q_stUps.LineInputVoltage_R := i_stState.fInputVoltageRV;
q_stUps.LineInputVoltage_S := i_stState.fInputVoltageSV;
q_stUps.LineInputVoltage_T := i_stState.fInputVoltageTV;
q_stUps.InputFrequency := i_stState.fInputFrequencyHz;
q_stUps.InputCurrent_R := i_stState.fInputCurrentRA;
q_stUps.InputCurrent_S := i_stState.fInputCurrentSA;
q_stUps.InputCurrent_T := i_stState.fInputCurrentTA;
q_stUps.InverterVoltage_R := i_stState.fInverterVoltageRV;
q_stUps.InverterVoltage_S := i_stState.fInverterVoltageSV;
q_stUps.InverterVoltage_T := i_stState.fInverterVoltageTV;
q_stUps.InverterCurrent_R := i_stState.fInverterCurrentRA;
q_stUps.InverterCurrent_S := i_stState.fInverterCurrentSA;
q_stUps.InverterCurrent_T := i_stState.fInverterCurrentTA;
q_stUps.BypassLineVoltage_R := i_stState.fBypassVoltageRV;
q_stUps.BypassLineVoltage_S := i_stState.fBypassVoltageSV;
q_stUps.BypassLineVoltage_T := i_stState.fBypassVoltageTV;
q_stUps.BypassFrequency := i_stState.fBypassFrequencyHz;
q_stUps.LineOutputVoltage_R := i_stState.fOutputVoltageRV;
q_stUps.LineOutputVoltage_S := i_stState.fOutputVoltageSV;
q_stUps.LineOutputVoltage_T := i_stState.fOutputVoltageTV;
q_stUps.FrequencyOutput := i_stState.fOutputFrequencyHz;
q_stUps.OutputCurrent_R := i_stState.fOutputCurrentRA;
q_stUps.OutputCurrent_S := i_stState.fOutputCurrentSA;
q_stUps.OutputCurrent_T := i_stState.fOutputCurrentTA;
q_stUps.DcLinkVoltage := i_stState.fDcLinkVoltageV;
q_stUps.DcLinkVoltage_High := i_stState.fDcLinkHighVoltageV;
q_stUps.DcLinkVoltage_Low := i_stState.fDcLinkLowVoltageV;
q_stUps.BatteryVoltage := i_stState.fBatteryVoltageV;
q_stUps.BatteryCurrent := i_stState.fBatteryCurrentA;
q_stUps.MPI_A_Current := i_stState.fMpiCurrentAA;
q_stUps.MPI_B_Current := i_stState.fMpiCurrentBA;
q_stUps.MPI_C_Current := i_stState.fMpiCurrentCA;
q_stUps.InputApparentPower := i_stState.fInputApparentPowerKva;
q_stUps.OutputApparentPower := i_stState.fOutputApparentPowerKva;
q_stUps.OutputActivePower := i_stState.fOutputActivePowerKw;
q_stUps.Temp1 := i_stState.fTemperature1C;
q_stUps.Temp2 := i_stState.fTemperature2C;
q_stUps.Temp3 := i_stState.fTemperature3C;
q_stUps.Temp4 := i_stState.fTemperature4C;
q_stUps.Temp5 := i_stState.fTemperature5C;
q_stUps.Temp6 := i_stState.fBatteryRoomTemperatureC;

END_FUNCTION_BLOCK

// ---- 20_Module/Report/FB_RptLsImd1000.TcPOU
FUNCTION_BLOCK FB_RptLsImd1000		// LS IMD1000 읽은 값 → IMD 보고값 (인터페이스\22. IMD.xlsx)
(* 2026-11-09. 명세 DV-11·RD-IMD-01 (v1.8)
   Status (사용자 결정 2026-11-09, 저항이 높은 경보부터)
     b0 통신에러 = 통신 이상 또는 아직 못 읽음 (나머지 칸 0)
     b1 Pre-Warning = Pre Alarm#3 동작 (IR 210 b3, 초기값 100 kΩ)
     b2 Warning = Pre Alarm#1 OR #2 동작 (IR 210 b1·b2, 초기값 40·70 kΩ)
     b3 Fault = 자가진단 오류 (IR 209 b0~2 메모리·RTC·교정) OR Device 이상 (IR 211 b1)
     b4 Alarm = Ins. Alarm 동작 (IR 210 b0, 초기값 10 kΩ)
     b5 Internal test = Self Test 진행 중 (IR 215 = 1)
     b6 External test = 버튼·DI Self Test 입력 (IR 206 b0·b1)
   Fault1 b0 = System 연결 이상 (IR 211 b2), b1 = PE 연결 이상 (IR 211 b0)
   PreAlarmSettingValue = Pre Alarm#1 Pick-up, MainAlarmSettingValue = Ins. Alarm Pick-up (설정 영역을 못 읽었으면 0)
   DeviceErrorLocation·InsulationResistanceFaultLocation은 Bender 항목이라 0 *)
VAR_INPUT
	i_stState		: ST_LsImd1000State;	// 장비 상태 (FB_LsImd1000.q_stState)
	i_nDeviceIndex	: UDINT;				// IMD 번호 (1부터)
END_VAR
VAR_OUTPUT
	q_stImd			: ST_ImdPublish_V1;		// IMD 보고값
	q_bValid		: BOOL;					// 유효한 장비 데이터
END_VAR
VAR
	_stEmpty		: ST_ImdPublish_V1;
END_VAR

q_stImd := _stEmpty;
q_stImd.DeviceIndex := i_nDeviceIndex;
q_stImd.Status := 1;	// b0 통신에러
q_bValid := i_stState.bValid;
IF NOT q_bValid THEN
	RETURN;
END_IF

q_stImd.Status := 0;
q_stImd.Status.1 := i_stState.wAlarm.3;
q_stImd.Status.2 := i_stState.wAlarm.1 OR i_stState.wAlarm.2;
q_stImd.Status.3 := (i_stState.wSelfDiag AND 16#0007) <> 0 OR i_stState.wConnect.1;
q_stImd.Status.4 := i_stState.wAlarm.0;
q_stImd.Status.5 := i_stState.wSelfTest = 1;
q_stImd.Status.6 := i_stState.wDiState.0 OR i_stState.wDiState.1;

q_stImd.InsulationResistance := i_stState.fInsulation;
IF i_stState.bSetValid THEN
	q_stImd.PreAlarmSettingValue := i_stState.nPre1Pickup;
	q_stImd.MainAlarmSettingValue := i_stState.nInsPickup;
END_IF
q_stImd.Fault1.0 := i_stState.wConnect.2;
q_stImd.Fault1.1 := i_stState.wConnect.0;

END_FUNCTION_BLOCK

// ---- 20_Module/Report/FB_RptTempHum.TcPOU
FUNCTION_BLOCK FB_RptTempHum		// 온습도계 읽은 값 → 온도 보고값 (인터페이스\07.Temperature Sensor.xlsx, 토픽 temperature_sensor)
(* 2026-11-09. status b0 통신에러(통신 이상·값 무효면 1, 온도·습도 0). location은 설치 위치 번호
   (1 PCS실, 2 BAT실, 3 UPS실, 4 FC 컨테이너실, 5 외부) *)
VAR_INPUT
	i_stState		: ST_TempHumState;		// 장비 상태 (드라이버 q_stState)
	i_nDeviceIndex	: UDINT;				// 장치 번호 (0부터, 기존 temperature_sensor 시험 데이터와 같음)
	i_nLocation		: UDINT;				// 설치 위치
END_VAR
VAR_OUTPUT
	q_stTemp		: ST_TempPublish_V1;	// 보고값
	q_bValid		: BOOL;					// 유효한 장비 데이터
END_VAR
VAR
	_stEmpty		: ST_TempPublish_V1;
END_VAR

q_stTemp := _stEmpty;
q_stTemp.DeviceIndex := i_nDeviceIndex;
q_stTemp.location := i_nLocation;
q_stTemp.status := 1;	// b0 통신에러
q_bValid := i_stState.bValid;
IF NOT q_bValid THEN
	RETURN;
END_IF
q_stTemp.status := 0;
q_stTemp.temperature := i_stState.fTemp;
q_stTemp.humidity := i_stState.fHum;

END_FUNCTION_BLOCK

// ---- 20_Module/Driver/Esolution/FB_BmsRackCommand.TcPOU
FUNCTION_BLOCK FB_BmsRackCommand		// BMS 랙 컨택터 개별 제어: EMS 랙 명령 → 랙 선택표(BMS 40001 랙 비트) 갱신 요청
(* 2026-11-10. 명세 WR-BAT-01 (v2.5). 인터페이스 100.Command BAT CommandType 11 랙 닫기 / 12 랙 열기 (Value = 랙 번호)
   BAT 질의 Q4 답변: 랙 개별·일괄 제어 모두 지원. 일괄은 CommandType 1·2 (시스템 컨택터 40013, 기존 코어 경로)
   - 랙 선택표(비트 n-1 = 랙 n, 1 = 사용)를 기억하고, 명령마다 그 랙 비트만 바꾼 표 전체를 BMS에 쓰게 한다
   - 장비 쓰기는 하지 않는다. q_bWriteReq·q_wWriteMask를 MAIN이 보고 드라이버 M_SetRackMask를 부르고 결과를 돌려준다
   - 선택표는 PERSISTENT (i_wRestore로 시작 때 한 번 읽고, q_wMask를 MAIN이 저장). 저장값이 없으면(0) 설치된 랙 전부
   - 거절: 랙 번호 범위 밖(BadRequest), 마지막 남은 랙 열기(BadRequest: 0이면 BMS가 전 랙 사용 안 함 → 전체는 일괄 2 열기로)
   - 드라이버가 바쁘면(Busy) WRITE_TIMEOUT 동안 다시 시도. 그 밖의 거절(쓰기 막힘, 통신 불가 등)은 바로 그 결과로 끝
   - 같은 상태로 바꾸는 명령도 표 전체를 다시 씀 (BMS가 다시 켜져 표가 달라졌을 때 맞춤)
   - [2026-11-13] BMS 맵 v1.4 랙 컨택터 상태(Input 30027)를 받으면 그 실제 상태를 바탕으로 비트를 바꿈.
     40013(랙 전체 연결)으로 다 붙은 뒤 옛 선택표로 써서 다른 랙을 떼는 일을 막음. 상태가 없으면 기억한 선택표 *)
VAR_INPUT
	i_stCmd			: ST_BatRackCmd;	// EMS 랙 명령 (번호가 바뀌면 새 명령)
	i_nRackCount	: UINT;				// 설치된 랙 수 (GVL_PARAM.RACKS_PER_BMS)
	i_wRestore		: WORD;				// 처음 호출 때 한 번 읽는 저장된 선택표 (GVL_PERSIST.g_awBmsRackMask[n])
	i_bAccepted		: BOOL;				// 지난 스캔의 쓰기 요청을 드라이버가 받음 (M_SetRackMask 반환값)
	i_eDriverResult	: E_UpsResult;		// 지난 스캔 드라이버 결과 (q_eRequestResult). 요청하지 않은 스캔은 None
	i_wActual		: WORD;				// BMS 랙 컨택터 실제 상태 (q_stState.wRackContactor, 30027) [2026-11-13]
	i_bActualValid	: BOOL;				// i_wActual을 믿을 수 있음 (q_stState.bContactorFeedbackKnown)
END_VAR
VAR_OUTPUT
	q_wMask			: WORD;				// 지금 선택표 (드라이버가 받은 값). MAIN이 GVL_PERSIST에 씀
	q_bMaskChanged	: BOOL;				// 이 스캔에 q_wMask가 바뀜 (PERSISTENT 바로 저장 요청)
	q_bWriteReq		: BOOL;				// 드라이버에 쓰기 요청 중
	q_wWriteMask	: WORD;				// 쓸 선택표
	q_eResult		: E_UpsResult;		// 마지막 명령 결과
	q_nLastSeq		: UDINT;			// 마지막으로 처리한 명령 번호
END_VAR
VAR
	_bInit			: BOOL;
	_wInstalled		: WORD;
	_wNew			: WORD;
	_wOld			: WORD;
	_wBase			: WORD;				// 바꿀 바탕 (실제 상태 또는 기억한 선택표)
	_tonWait		: TON;
END_VAR
VAR CONSTANT
	WRITE_TIMEOUT	: TIME := T#5S;		// 드라이버가 바쁠 때 다시 시도하는 시간
END_VAR

q_bMaskChanged := FALSE;
_wInstalled := SHL(WORD#1, MIN(i_nRackCount, 16)) - 1;
IF NOT _bInit THEN
	q_wMask := i_wRestore AND _wInstalled;
	IF q_wMask = 0 THEN
		q_wMask := _wInstalled;	// 저장값 없음 → 설치된 랙 전부
	END_IF
	_bInit := TRUE;
END_IF
_wOld := q_wMask;

// 1) 지난 스캔 쓰기 요청의 결과
IF q_bWriteReq THEN
	_tonWait(IN := TRUE, PT := WRITE_TIMEOUT);
	IF i_bAccepted THEN
		q_wMask := q_wWriteMask;
		q_eResult := E_UpsResult.Accepted;
		q_bWriteReq := FALSE;
	ELSIF i_eDriverResult <> E_UpsResult.None AND i_eDriverResult <> E_UpsResult.Busy THEN
		q_eResult := i_eDriverResult;	// 쓰기 막힘, 통신 불가, 설정 오류 등
		q_bWriteReq := FALSE;
	ELSIF _tonWait.Q THEN
		q_eResult := E_UpsResult.Busy;	// 계속 바빠서 포기
		q_bWriteReq := FALSE;
	END_IF
	IF NOT q_bWriteReq THEN
		_tonWait(IN := FALSE);
	END_IF
END_IF

// 2) 새 명령 (처리 중인 요청이 있으면 그것을 버리고 새 명령으로)
IF i_stCmd.nSeq <> q_nLastSeq AND i_stCmd.nSeq <> 0 THEN
	q_nLastSeq := i_stCmd.nSeq;
	q_bWriteReq := FALSE;
	_tonWait(IN := FALSE);
	IF i_stCmd.nRack < 1 OR i_stCmd.nRack > i_nRackCount OR i_stCmd.nRack > 16 THEN
		q_eResult := E_UpsResult.BadRequest;
	ELSE
		IF i_bActualValid THEN
			_wBase := i_wActual AND _wInstalled;	// 실제 상태 바탕
		ELSE
			_wBase := q_wMask;
		END_IF
		IF i_stCmd.bClose THEN
			_wNew := _wBase OR SHL(WORD#1, i_stCmd.nRack - 1);
		ELSE
			_wNew := _wBase AND NOT SHL(WORD#1, i_stCmd.nRack - 1);
		END_IF
		IF _wNew = 0 THEN
			q_eResult := E_UpsResult.BadRequest;	// 마지막 랙: 전체 열기는 일괄 명령(2)으로
		ELSE
			q_wWriteMask := _wNew;
			q_bWriteReq := TRUE;
			q_eResult := E_UpsResult.None;	// 처리 중
		END_IF
	END_IF
END_IF

q_bMaskChanged := q_wMask <> _wOld;

END_FUNCTION_BLOCK

// ---- 20_Module/Driver/Esolution/FB_BmsContactorCommand.TcPOU
FUNCTION_BLOCK FB_BmsContactorCommand		// BMS 컨택터 하나씩 제어: EMS 명령 번호 5~10 → 드라이버 M_SetControl 요청
(* 2026-11-13. 인터페이스 100.Command BAT CommandType 5~10, BMS 맵 v1.4 Holding 40013~40015
   5 시스템(랙 전체 40013) 연결   6 시스템 차단
   7 충전 컨택터(40014) 닫기      8 충전 컨택터 열기
   9 방전 컨택터(40015) 닫기      10 방전 컨택터 열기
   - 장비 쓰기는 하지 않는다. q_bWriteReq·q_eControl·q_bOn을 MAIN이 보고 드라이버 M_SetControl을 부르고 결과를 돌려준다
   - 5~10 밖이면 BadRequest. 드라이버가 바쁘면(Busy) WRITE_TIMEOUT 동안 다시 시도. 그 밖의 거절(쓰기 막힘, 통신 불가 등)은 바로 그 결과로 끝
   - 코어 순서(유닛 정지 확인)는 거치지 않는다 (랙 개별 11·12와 같음). 일괄 투입·개방은 1·2 (코어 경로) *)
VAR_INPUT
	i_stCmd			: ST_BatCtlCmd;		// EMS 명령 (번호가 바뀌면 새 명령)
	i_bAccepted		: BOOL;				// 지난 스캔의 쓰기 요청을 드라이버가 받음 (M_SetControl 반환값)
	i_eDriverResult	: E_UpsResult;		// 지난 스캔 드라이버 결과 (q_eRequestResult). 요청하지 않은 스캔은 None
END_VAR
VAR_OUTPUT
	q_bWriteReq		: BOOL;				// 드라이버에 쓰기 요청 중
	q_eControl		: E_EsolutionControl;	// 쓸 컨택터
	q_bOn			: BOOL;				// TRUE = 닫기(붙이기), FALSE = 열기(떼기)
	q_eResult		: E_UpsResult;		// 마지막 명령 결과
	q_nLastSeq		: UDINT;			// 마지막으로 처리한 명령 번호
END_VAR
VAR
	_tonWait		: TON;
END_VAR
VAR CONSTANT
	WRITE_TIMEOUT	: TIME := T#5S;		// 드라이버가 바쁠 때 다시 시도하는 시간
END_VAR

// 1) 지난 스캔 쓰기 요청의 결과
IF q_bWriteReq THEN
	_tonWait(IN := TRUE, PT := WRITE_TIMEOUT);
	IF i_bAccepted THEN
		q_eResult := E_UpsResult.Accepted;
		q_bWriteReq := FALSE;
	ELSIF i_eDriverResult <> E_UpsResult.None AND i_eDriverResult <> E_UpsResult.Busy THEN
		q_eResult := i_eDriverResult;	// 쓰기 막힘, 통신 불가 등
		q_bWriteReq := FALSE;
	ELSIF _tonWait.Q THEN
		q_eResult := E_UpsResult.Busy;	// 계속 바빠서 포기
		q_bWriteReq := FALSE;
	END_IF
	IF NOT q_bWriteReq THEN
		_tonWait(IN := FALSE);
	END_IF
END_IF

// 2) 새 명령 (처리 중인 요청이 있으면 그것을 버리고 새 명령으로)
IF i_stCmd.nSeq <> q_nLastSeq AND i_stCmd.nSeq <> 0 THEN
	q_nLastSeq := i_stCmd.nSeq;
	q_bWriteReq := FALSE;
	_tonWait(IN := FALSE);
	q_eResult := E_UpsResult.None;	// 처리 중
	CASE i_stCmd.nType OF
		5, 6:	q_eControl := E_EsolutionControl.SystemContactor;
		7, 8:	q_eControl := E_EsolutionControl.ChargeContactor;
		9, 10:	q_eControl := E_EsolutionControl.DischargeContactor;
	ELSE
		q_eResult := E_UpsResult.BadRequest;
	END_CASE
	IF q_eResult = E_UpsResult.None THEN
		q_bOn := (i_stCmd.nType MOD 2) = 1;	// 5·7·9 = 닫기
		q_bWriteReq := TRUE;
	END_IF
END_IF

END_FUNCTION_BLOCK

// ---- 20_Module/Ups/FB_UpsSafetyStage.TcPOU
(* LiB-UPS 사고·고장 단계 판정 (④보호 표시 / 장치: UPS·BAT). 2026-11-05.
   기반 없음(신규). 동작시퀀스 7쪽(이솔루션 2026-10-23) 단계표를 따른다.
   변경: 2026-11-09 UPS 경고·고장 4번 칸을 없앰. STATUS 비트를 Warning3 하위·Fault3 상위에서 읽음 (명세 RD-UPS-02 v1.6)
   부호·단위: 해당 없음. 명세: C:\gil\UPS\명세서\UPS_명세서.md SQ-01, WR-SQ-01
   차단·정지는 UPS(UMS)와 BMS가 스스로 한다. 이 FB는 판정과 표시만 하고 장비에 아무것도 쓰지 않는다. *)
FUNCTION_BLOCK FB_UpsSafetyStage
VAR_INPUT
	i_stUps			: ST_UpsPublish_V1;	// UPS 보고값 (FB_RptSebangUps.q_stUps)
	i_bUpsValid		: BOOL;				// UPS 데이터 유효 (통신 정상)
	i_stBat			: ST_BatPublish_V1;	// 짝 BAT 보고값 (FB_RptEsolutionBat.q_stBat)
	i_bBatValid		: BOOL;				// BAT 데이터 유효 (통신 정상)
	i_bAck			: BOOL;				// Fault 단계 확인 (상승 에지). 원인이 해소된 Fault 표시만 내린다 (WR-SQ-01)
END_VAR
VAR_OUTPUT
	q_nStage		: UINT;				// 대표 단계 0~6 (걸린 단계 중 가장 높은 것)
	q_wStageMask	: WORD;				// 걸린 단계 목록. bit n = n단계 (n = 1~6). 높은 순서로 모두 표시할 때 사용
	q_nCause		: UDINT;			// 원인 비트 (아래 CAUSE_* 표). 지금 걸린 원인 + 확인 전인 Fault 원인
	q_nActiveCause	: UDINT;			// 지금 실제로 걸린 원인만
	q_bAckPending	: BOOL;				// 원인은 해소됐지만 운영자 확인 전인 Fault 원인이 있음
	q_bUpsCommFault	: BOOL;				// UPS 통신장애 (단계와 별도 상태). 끊긴 동안 UPS 원인은 마지막 값을 유지
	q_bBatCommFault	: BOOL;				// BAT 통신장애 (단계와 별도 상태). 끊긴 동안 BAT 원인은 마지막 값을 유지
END_VAR
VAR
	_rtAck			: R_TRIG;
	_nUpsCause		: UDINT;			// UPS에서 나온 원인 (통신이 끊기면 마지막 값 유지)
	_nBatCause		: UDINT;			// BAT에서 나온 원인 (통신이 끊기면 마지막 값 유지)
	_nLatched		: UDINT;			// 확인 전까지 유지하는 Fault 원인
	_i				: INT;
END_VAR
VAR CONSTANT
	(* 원인 비트 → 단계. 순서 = 비트 번호 *)
	CAUSE_STAGE		: ARRAY[0..12] OF UINT := [
		1,	// b0  AC·DC SPD (I51 b8·b9)
		1,	// b1  UPS 경고장 (SPD·BMS Minor 제외)
		2,	// b2  BMS Minor (I51 b10)
		3,	// b3  BMS Major (I51 b11)
		3,	// b4  UPS 입력·정류부 중고장 (Fault1)
		3,	// b5  UPS 출력 중고장 (Fault2 상위)
		3,	// b6  UPS 인버터 중고장 (Fault3 하위)
		3,	// b7  배터리 DC 전로 지락 1단계 = RCD 1단계 (I51 b12, 추정)
		4,	// b8  배터리 컨버터(BBC) 중고장 (Fault2 하위)
		4,	// b9  지락 2단계 = RCD 2단계 (I51 b13, 추정)
		5,	// b10 BMS Level 3 (BAT Status b9 System Lock)
		5,	// b11 화재 (I51 b14)
		6];	// b12 ESD (I50 b0)
	FAULT_CAUSE_MASK : UDINT := 16#00001F00;	// 4~6단계 원인 (b8~b12): 확인 전까지 유지
	(* UPS 보고 칸 안의 비트 (명세 RD-UPS-02 v1.6). Warning3 하위 16비트 = I51 경고, Fault3 상위 16비트 = I50 고장 OR I51 고장 *)
	W3_SPD			: UDINT := 16#00000300;	// Warning3: I51 b8 AC SPD, b9 DC SPD
	W3_BMS_MINOR	: UDINT := 16#00000400;	// Warning3: I51 b10
	F3_BMS_MAJOR	: UDINT := 16#08000000;	// Fault3: I51 b11
	F3_RCD1			: UDINT := 16#10000000;	// Fault3: I51 b12
	F3_RCD2			: UDINT := 16#20000000;	// Fault3: I51 b13
	F3_FIRE			: UDINT := 16#40000000;	// Fault3: I51 b14
	F3_ESD			: UDINT := 16#00010000;	// Fault3: I50 b0
	LOWER_WORD		: UDINT := 16#0000FFFF;
	UPPER_WORD		: UDINT := 16#FFFF0000;
END_VAR

// 1) UPS 원인. 통신이 끊기면 마지막 값을 그대로 둔다 (단계를 내리지 않음)
q_bUpsCommFault := NOT i_bUpsValid;
IF i_bUpsValid THEN
	_nUpsCause := 0;
	IF (i_stUps.Warning3 AND W3_SPD) <> 0 THEN _nUpsCause := _nUpsCause OR 16#0001; END_IF
	IF (i_stUps.Warning1 OR i_stUps.Warning2 OR (i_stUps.Warning3 AND NOT (W3_SPD OR W3_BMS_MINOR))) <> 0 THEN _nUpsCause := _nUpsCause OR 16#0002; END_IF
	IF (i_stUps.Warning3 AND W3_BMS_MINOR) <> 0 THEN _nUpsCause := _nUpsCause OR 16#0004; END_IF
	IF (i_stUps.Fault3 AND F3_BMS_MAJOR) <> 0 THEN _nUpsCause := _nUpsCause OR 16#0008; END_IF
	IF i_stUps.Fault1 <> 0 THEN _nUpsCause := _nUpsCause OR 16#0010; END_IF
	IF (i_stUps.Fault2 AND UPPER_WORD) <> 0 THEN _nUpsCause := _nUpsCause OR 16#0020; END_IF
	IF (i_stUps.Fault3 AND LOWER_WORD) <> 0 THEN _nUpsCause := _nUpsCause OR 16#0040; END_IF
	IF (i_stUps.Fault3 AND F3_RCD1) <> 0 THEN _nUpsCause := _nUpsCause OR 16#0080; END_IF
	IF (i_stUps.Fault2 AND LOWER_WORD) <> 0 THEN _nUpsCause := _nUpsCause OR 16#0100; END_IF
	IF (i_stUps.Fault3 AND F3_RCD2) <> 0 THEN _nUpsCause := _nUpsCause OR 16#0200; END_IF
	IF (i_stUps.Fault3 AND F3_FIRE) <> 0 THEN _nUpsCause := _nUpsCause OR 16#0800; END_IF
	IF (i_stUps.Fault3 AND F3_ESD) <> 0 THEN _nUpsCause := _nUpsCause OR 16#1000; END_IF
END_IF

// 2) BAT 원인
q_bBatCommFault := NOT i_bBatValid;
IF i_bBatValid THEN
	_nBatCause := 0;
	IF i_stBat.Status.9 THEN _nBatCause := _nBatCause OR 16#0400; END_IF	// BMS Level 3 (System Lock)
END_IF

q_nActiveCause := _nUpsCause OR _nBatCause;

// 3) Fault(4~6단계)는 원인이 사라져도 확인 전까지 유지. 확인하면 해소된 것만 내림
_nLatched := _nLatched OR (q_nActiveCause AND FAULT_CAUSE_MASK);
_rtAck(CLK := i_bAck);
IF _rtAck.Q THEN
	_nLatched := _nLatched AND q_nActiveCause;
END_IF
q_nCause := q_nActiveCause OR _nLatched;
q_bAckPending := (_nLatched AND NOT q_nActiveCause) <> 0;

// 4) 단계 목록과 대표 단계
q_wStageMask := 0;
q_nStage := 0;
FOR _i := 0 TO 12 DO
	IF (q_nCause AND SHL(UDINT#1, _i)) <> 0 THEN
		q_wStageMask := q_wStageMask OR SHL(WORD#1, CAUSE_STAGE[_i]);
		q_nStage := MAX(q_nStage, CAUSE_STAGE[_i]);
	END_IF
END_FOR

END_FUNCTION_BLOCK

// ---- 20_Module/Mqtt/FB_EmsConfigApply.TcPOU
FUNCTION_BLOCK FB_EmsConfigApply		// EMS config(pcs·bat) → 운영 설정 (PlcTask. MAIN 액션 A_PassEmsCfg가 부름) [9-21 수정 2026-11-04: 추가]
(* - 입력 i_stCfg는 MAIN이 GVL_IF.g_stEmsCfg에서 일관되게 복사해 넘김. PCS·BMS 칸마다 번호(anPcsSeq·anBatSeq)가 바뀌면 새 레코드
   - [21번 수정 2026-11-09] is_available = 0인 값은 기본값으로 반영 (원래: 바꾸지 않고 기존 값 유지 → EMS가 한도를 풀 수 없었음)
       pcs 충전·방전 한도 0 → 그 방향 정격 (= 제한 없음). 두 방향 모두 0 → 그 PCS 유닛의 사용자 P 한도 끔 (bPEnable FALSE, 값은 ±정격)
       bat SOC 하한 0 → 0 %, 상한 0 → 100 % (감발 폭 fBand·재개 마진은 HMI 설정 그대로)
   - [UPS 2026-11-10] UPS 현장의 config/bat 레코드는 103.Config BAT UPS_V1 형식 (SocMin·SocMax = REAL, is_available 없음. UPS_MQTT_INTERFACE.md).
       그래서 bat 값은 받은 BMS(_abBatRx)만 계산에 넣고 항상 '있음'으로 봄. 아직 못 받은 BMS는 기본값(0 %·100 %)과 같아 결과에 영향 없음. pcs 쪽은 STD 그대로
   - pcs: 충전·방전 전력 한도 (kW) → 사용자 한도 stUnitLimit. 그 PCS의 유닛들에 정격 비율로 나눔, 충전은 fPMin (−). PvMarginRate는 쓰지 않음 (사양 대기)
   - bat: SOC 최소·최대 (%) → SOC 정책 stSocLimit. 배터리 그룹 전체 한 세트라 받은 BMS 값(기본값 포함) 중 가장 엄격한 값 (하한 = 가장 큰 값, 상한 = 가장 작은 값)
   - 범위 검사를 먼저 하고 통과한 값만 씀 (SOC는 FB_SocLimit.M_CheckSet과 같은 F_SocLimitSetErr). 버리면 q_bRejected (이벤트 로그 '잘못된 설정 값')
   - 쓴 값은 GVL_PERSIST라 재시작 뒤에도 남음. 설정 보호(FB_SettingGuard)가 한 번 더 지킴. 바꾸면 q_bApplied (이벤트 로그 '운영 설정 바뀜')
   - protection(배터리·배터리실 온도·습도 경고·고장)은 반영하지 않음 (값의 뜻·센서 대기. echo만)
   - M_BuildEcho: 설정 보호 뒤 실제 설정 → q_stEcho (MAIN이 GVL_IF.g_stEmsCfgEcho에 씀 → config echo) *)
VAR_INPUT
	i_bValid		: BOOL;			// 이번 스캔에 i_stCfg를 일관되게 복사함
	i_stCfg			: ST_IfEmsCfg;
	i_astUnitCfg	: ARRAY[1..GVL_PARAM.UNIT_COUNT] OF ST_UnitCfg;	// 유닛 ← PCS 번호, 정격
END_VAR
VAR_IN_OUT
	iq_stSocLimit	: ST_SocLimitSet;	// GVL_PERSIST.g_stModuleSet.stSocLimit
	iq_stUnitLimit	: ST_UnitLimitSet;	// GVL_PERSIST.g_stModuleSet.stUnitLimit
END_VAR
VAR_OUTPUT
	q_bApplied		: BOOL;			// 이번 스캔에 설정을 바꿈 (1스캔)
	q_sApplied		: WSTRING(63);
	q_bRejected		: BOOL;			// 이번 스캔에 받은 값을 버림 (1스캔)
	q_sRejected		: WSTRING(63);	// 마지막으로 버린 값과 이유
	q_nApplied		: UDINT;
	q_nRejected		: UDINT;
	q_stEcho		: ST_IfEmsCfgEcho;
END_VAR
VAR CONSTANT
	MAX_KW			: REAL := 1.0E6;	// kW. 이보다 큰 한도는 이상값
	SOC_MIN_DEFAULT	: REAL := 0.0;		// %, bat SocMin is_available 0일 때 [21번 수정 2026-11-09: 추가]
	SOC_MAX_DEFAULT	: REAL := 100.0;	// %, bat SocMax is_available 0일 때
END_VAR
VAR
	_stCfg			: ST_IfEmsCfg;		// 마지막으로 일관되게 받은 칸 (echo의 PvMarginRate)
	_anPcsSeq		: ARRAY[1..GVL_PARAM.PCS_COUNT] OF UDINT;
	_anBatSeq		: ARRAY[1..GVL_PARAM.BMS_COUNT] OF UDINT;
	_astBat			: ARRAY[1..GVL_PARAM.BMS_COUNT] OF ST_BatConfig_Rx;	// BMS마다 받아 둔 레코드 (가장 엄격한 SOC 계산)
	_astBatBefore	: ARRAY[1..GVL_PARAM.BMS_COUNT] OF ST_BatConfig_Rx;
	_abBatRx		: ARRAY[1..GVL_PARAM.BMS_COUNT] OF BOOL;	// [UPS] 그 BMS 레코드를 한 번이라도 받아 둠 (REAL 형식이라 빈 칸을 is_available로 못 가림)
	_abBatRxBefore	: ARRAY[1..GVL_PARAM.BMS_COUNT] OF BOOL;
	_stUnit			: ST_UnitLimitSet;
	_stSoc			: ST_SocLimitSet;
	_sErr			: WSTRING(63);
	p				: UINT;
	u				: UINT;
	b				: UINT;
	fSum			: REAL;
	fCh				: REAL;
	fDis			: REAL;
	fMin			: REAL;
	fMax			: REAL;
	bCh				: BOOL;
	bDis			: BOOL;
	bAny			: BOOL;
	bNewBat			: BOOL;
	bBad			: BOOL;
END_VAR

q_bApplied	:= FALSE;
q_bRejected	:= FALSE;
IF NOT i_bValid THEN
	RETURN;
END_IF
_stCfg := i_stCfg;

(* PCS: 충전·방전 전력 한도 → 그 PCS 유닛들의 사용자 한도 (정격 비율) *)
_stUnit := iq_stUnitLimit;
bAny := FALSE;
FOR p := 1 TO GVL_PARAM.PCS_COUNT DO
	IF i_stCfg.anPcsSeq[p] <> _anPcsSeq[p] THEN
		_anPcsSeq[p] := i_stCfg.anPcsSeq[p];
		bCh		:= i_stCfg.astPcs[p].ChargePowerLimit.is_available <> 0;
		bDis	:= i_stCfg.astPcs[p].DisChargePowerLimit.is_available <> 0;
		fCh		:= UDINT_TO_REAL(i_stCfg.astPcs[p].ChargePowerLimit.value);
		fDis	:= UDINT_TO_REAL(i_stCfg.astPcs[p].DisChargePowerLimit.value);
		fSum := 0.0;
		FOR u := 1 TO GVL_PARAM.UNIT_COUNT DO
			IF i_astUnitCfg[u].nPcs = p AND F_RealOk(i_astUnitCfg[u].fPRated) THEN
				fSum := fSum + i_astUnitCfg[u].fPRated;
			END_IF
		END_FOR
		IF (bCh AND fCh > MAX_KW) OR (bDis AND fDis > MAX_KW) THEN
			M_Reject(F_TxtNum("EMS config pcs 전력 한도 범위 밖: PCS ", p));
		ELSIF NOT (fSum > 0.0) THEN
			M_Reject(F_TxtNum("EMS config pcs 유닛 없음(정격 합 0): PCS ", p));
		ELSE
			// [21번 수정 2026-11-09: is_available 0인 방향은 정격(제한 없음), 둘 다 0이면 사용자 P 한도 끔.
			//   원래: 둘 다 0이면 아무것도 안 바꿈, 한쪽만 0이면 그 방향은 기존 값 유지 (처음 켤 때만 정격)]
			FOR u := 1 TO GVL_PARAM.UNIT_COUNT DO
				IF i_astUnitCfg[u].nPcs = p THEN
					_stUnit.astUnit[u].bPEnable	:= bCh OR bDis;
					IF bDis THEN
						_stUnit.astUnit[u].fPMax := fDis * MAX(i_astUnitCfg[u].fPRated, 0.0) / fSum;
					ELSE
						_stUnit.astUnit[u].fPMax := MAX(i_astUnitCfg[u].fPRated, 0.0);
					END_IF
					IF bCh THEN
						_stUnit.astUnit[u].fPMin := -(fCh * MAX(i_astUnitCfg[u].fPRated, 0.0) / fSum);
					ELSE
						_stUnit.astUnit[u].fPMin := -MAX(i_astUnitCfg[u].fPRated, 0.0);
					END_IF
				END_IF
			END_FOR
			bAny := TRUE;
		END_IF
	END_IF
END_FOR
IF bAny AND MEMCMP(ADR(_stUnit), ADR(iq_stUnitLimit), SIZEOF(_stUnit)) <> 0 THEN
	iq_stUnitLimit := _stUnit;
	M_Applied("EMS config: PCS 충·방전 전력 한도");
END_IF

(* BMS: SOC 최소·최대 → SOC 정책 (가장 엄격한 값). 값마다 숫자·0~100 먼저, 합친 설정은 F_SocLimitSetErr *)
_astBatBefore := _astBat;
_abBatRxBefore := _abBatRx;
bNewBat := FALSE;
FOR b := 1 TO GVL_PARAM.BMS_COUNT DO
	IF i_stCfg.anBatSeq[b] <> _anBatSeq[b] THEN
		_anBatSeq[b] := i_stCfg.anBatSeq[b];
		bBad := FALSE;
		// [UPS] SocMin·SocMax는 REAL (is_available 없음) → 둘 다 항상 검사
		bBad := NOT (F_RealOk(i_stCfg.astBat[b].SocMin) AND_THEN (i_stCfg.astBat[b].SocMin >= 0.0 AND i_stCfg.astBat[b].SocMin <= 100.0));
		IF NOT bBad THEN
			bBad := NOT (F_RealOk(i_stCfg.astBat[b].SocMax) AND_THEN (i_stCfg.astBat[b].SocMax >= 0.0 AND i_stCfg.astBat[b].SocMax <= 100.0));
		END_IF
		IF bBad THEN
			M_Reject(F_TxtNum("EMS config bat SOC 숫자·범위(0~100) 아님: BMS ", b));
		ELSE
			_astBat[b] := i_stCfg.astBat[b];
			_abBatRx[b] := TRUE;
			bNewBat := TRUE;
		END_IF
	END_IF
END_FOR
IF bNewBat THEN
	// [21번 수정 2026-11-09: is_available 0이면 기본값(하한 0 %, 상한 100 %)으로 보고 가장 엄격한 값을 고름. 기본값은 다른 BMS 값보다 엄격하지 않으므로
	//   값을 하나도 안 받은 BMS(빈 칸)는 결과에 영향이 없음. 원래: is_available 0은 계산에서 빼고, 하나도 없으면 기존 값 유지]
	fMin := SOC_MIN_DEFAULT;
	fMax := SOC_MAX_DEFAULT;
	FOR b := 1 TO GVL_PARAM.BMS_COUNT DO
		IF _abBatRx[b] AND_THEN _astBat[b].SocMin > fMin THEN		// [UPS] 받은 BMS만 (원래 SocMin.is_available <> 0 AND_THEN SocMin.value > fMin)
			fMin := _astBat[b].SocMin;
		END_IF
		IF _abBatRx[b] AND_THEN _astBat[b].SocMax < fMax THEN
			fMax := _astBat[b].SocMax;
		END_IF
	END_FOR
	_stSoc := iq_stSocLimit;
	_stSoc.fSocMin := fMin;
	_stSoc.fSocMax := fMax;
	_sErr := F_SocLimitSetErr(_stSoc);
	IF _sErr <> "" THEN
		_astBat := _astBatBefore;		// 이번에 받은 BMS 값은 버림 (다음 계산에 쓰지 않음)
		_abBatRx := _abBatRxBefore;
		M_Reject(WCONCAT("EMS config bat: ", _sErr));
	ELSIF MEMCMP(ADR(_stSoc), ADR(iq_stSocLimit), SIZEOF(_stSoc)) <> 0 THEN
		iq_stSocLimit := _stSoc;
		M_Applied("EMS config: SOC 상·하한");
	END_IF
END_IF

METHOD PRIVATE M_Reject
VAR_INPUT
	i_sText	: WSTRING(63);
END_VAR
q_bRejected	:= TRUE;
q_sRejected	:= i_sText;
q_nRejected	:= q_nRejected + 1;
END_METHOD

METHOD PRIVATE M_Applied
VAR_INPUT
	i_sText	: WSTRING(63);
END_VAR
q_bApplied	:= TRUE;
q_sApplied	:= i_sText;
q_nApplied	:= q_nApplied + 1;
END_METHOD

METHOD M_BuildEcho		// 실제 설정 → q_stEcho (MAIN이 설정 보호 뒤에 부름)
VAR_IN_OUT CONSTANT
	iq_stSocLimit	: ST_SocLimitSet;
	iq_stUnitLimit	: ST_UnitLimitSet;
END_VAR
VAR
	p			: UINT;
	u			: UINT;
	b			: UINT;
	bAll		: BOOL;
	bUnit		: BOOL;
	fMaxSum		: REAL;
	fMinSum		: REAL;
END_VAR
FOR p := 1 TO GVL_PARAM.PCS_COUNT DO
	bAll	:= TRUE;
	bUnit	:= FALSE;
	fMaxSum	:= 0.0;
	fMinSum	:= 0.0;
	FOR u := 1 TO GVL_PARAM.UNIT_COUNT DO
		IF i_astUnitCfg[u].nPcs = p THEN
			bUnit := TRUE;
			IF iq_stUnitLimit.astUnit[u].bPEnable AND F_RealOk(iq_stUnitLimit.astUnit[u].fPMax) AND F_RealOk(iq_stUnitLimit.astUnit[u].fPMin) THEN
				fMaxSum := fMaxSum + iq_stUnitLimit.astUnit[u].fPMax;
				fMinSum := fMinSum + iq_stUnitLimit.astUnit[u].fPMin;
			ELSE
				bAll := FALSE;
			END_IF
		END_IF
	END_FOR
	q_stEcho.astPcs[p - 1].DeviceId := UINT_TO_UDINT(p);	// 번호 1부터 [1부터 2026-11-10]
	IF bUnit AND bAll THEN
		q_stEcho.astPcs[p - 1].DisChargePowerLimit.value		:= DINT_TO_UDINT(MAX(F_RealToDint(fMaxSum), 0));
		q_stEcho.astPcs[p - 1].DisChargePowerLimit.is_available	:= 1;
		q_stEcho.astPcs[p - 1].ChargePowerLimit.value			:= DINT_TO_UDINT(MAX(F_RealToDint(-fMinSum), 0));
		q_stEcho.astPcs[p - 1].ChargePowerLimit.is_available		:= 1;
	ELSE
		q_stEcho.astPcs[p - 1].DisChargePowerLimit.value		:= 0;
		q_stEcho.astPcs[p - 1].DisChargePowerLimit.is_available	:= 0;
		q_stEcho.astPcs[p - 1].ChargePowerLimit.value			:= 0;
		q_stEcho.astPcs[p - 1].ChargePowerLimit.is_available		:= 0;
	END_IF
	q_stEcho.astPcs[p - 1].PvMarginRate.value			:= _stCfg.astPcs[p].PvMarginRate.value;	// 쓰지 않음: 받은 값, is_available 0
	q_stEcho.astPcs[p - 1].PvMarginRate.is_available	:= 0;
END_FOR
FOR b := 1 TO GVL_PARAM.BMS_COUNT DO
	q_stEcho.astBat[b - 1].DeviceId					:= UINT_TO_UDINT(b);	// 번호 1부터 [1부터 2026-11-10]
	q_stEcho.astBat[b - 1].SocMin					:= iq_stSocLimit.fSocMin;	// [UPS] REAL 형식 (원래 SocMin.value + is_available 1)
	q_stEcho.astBat[b - 1].SocMax					:= iq_stSocLimit.fSocMax;
END_FOR
END_METHOD

END_FUNCTION_BLOCK

// ---- 20_Module/Common/F_SocLimitSetErr.TcPOU
FUNCTION F_SocLimitSetErr : WSTRING(63)		// SOC 정책 설정 점검 ("" = 정상). FB_SocLimit.M_CheckSet과 FB_EmsConfigApply(EMS config 반영 전 검사)가 같이 씀 [9-21 수정 2026-11-04: FB_SocLimit.M_CheckSet에서 옮김]
VAR_INPUT
	i_stSet	: ST_SocLimitSet;
END_VAR

F_SocLimitSetErr := "";
IF NOT (F_RealOk(i_stSet.fSocMin) AND F_RealOk(i_stSet.fSocMax) AND F_RealOk(i_stSet.fBand) AND F_RealOk(i_stSet.fResumeMargin)) THEN	// [결함 13 수정 2026-11-04]
	F_SocLimitSetErr := "SOC 설정 숫자 아님";
ELSIF i_stSet.fSocMin < 0.0 OR i_stSet.fSocMax > 100.0 OR i_stSet.fSocMin >= i_stSet.fSocMax THEN
	F_SocLimitSetErr := "SOC 상·하한 (0 ≤ 하한 < 상한 ≤ 100)";
ELSIF i_stSet.fBand < 0.0 OR i_stSet.fSocMin + i_stSet.fBand > i_stSet.fSocMax - i_stSet.fBand THEN
	F_SocLimitSetErr := "감발 폭 fBand (0 이상, 상·하한 사이)";
ELSIF i_stSet.fResumeMargin < 0.0 OR i_stSet.fSocMin + i_stSet.fResumeMargin >= i_stSet.fSocMax - i_stSet.fResumeMargin THEN
	F_SocLimitSetErr := "재개 마진 fResumeMargin (0 이상, 상·하한 사이)";
END_IF

END_FUNCTION

// ---- 20_Module/Mqtt/FB_BrokerWatch.TcPOU
FUNCTION_BLOCK FB_BrokerWatch		// MQTT 브로커 끊김 감시 (PlcTask, MAIN이 부름) [9번 수정 2026-11-09: 추가 — 14번 탭 9번 결정]
// - 감시: i_stSet.eBroker로 고른 브로커가 쓰는 브로커(MQTT_SET bUse)일 때만. 접속 상태는 PRG_Mqtt가 GVL_IF.g_abBrokerConn에 올림 (구독 클라이언트 기준)
// - 끊김: 접속이 i_stSet.tLostDelay 넘게 이어서 끊기면 q_bLost (알람 '브로커 끊김', 접속하면 해소). PMS 시작 직후 접속 전도 끊김으로 셈
// - Manual 전환: 끊김 동안 한 번만 q_bToManual (1스캔) → MAIN이 운전 모드 요청(g_aeOpMode)을 모두 Manual로. 끊긴 동안 운전원이 Auto로 되돌려도 다시 바꾸지 않음.
//   다시 접속하면(q_bLost 해소) 다시 무장 → 다음 끊김에 다시 한 번
// - 이중화: Active PLC만 전환 요청 (대기 PLC의 운전 모드 요청은 Active 값으로 동기화됨). 끊긴 동안 Active가 되면 그때 한 번
VAR_INPUT
	i_stSet			: ST_BrokerWatchSet;
	i_abUse			: ARRAY[1..3] OF BOOL;	// 쓰는 브로커 (GVL_IF.g_abBrokerUse, 1 Cloud, 2 Local, 3 Azure)
	i_abConnected	: ARRAY[1..3] OF BOOL;	// 접속됨 (GVL_IF.g_abBrokerConn)
	i_bActive		: BOOL;					// 이 PLC가 Active (GVL_IF.g_bRedActive. 이중화를 안 쓰면 항상 TRUE)
END_VAR
VAR_OUTPUT
	q_bWatch		: BOOL;			// 감시 중 (고른 브로커를 씀)
	q_bLost			: BOOL;			// 끊김 확정 (알람)
	q_bToManual		: BOOL;			// 이번 스캔에 Manual 전환 요청 (1스캔)
	q_sBroker		: WSTRING(15);	// 고른 브로커 이름 (로그)
	q_sDelay		: WSTRING(31);	// 판정 시간 글자 (로그)
END_VAR
VAR
	_tonLost		: TON;
	_bDone			: BOOL;			// 이번 끊김에서 전환 요청을 냄 (접속하면 지움)
	_n				: INT;			// 고른 브로커 칸 (0 = 범위 밖)
END_VAR

CASE i_stSet.eBroker OF
	E_MqttBroker.Cloud:	_n := 1;	q_sBroker := "Cloud";
	E_MqttBroker.Local:	_n := 2;	q_sBroker := "Local";
	E_MqttBroker.Azure:	_n := 3;	q_sBroker := "Azure";
ELSE
	_n := 0;	q_sBroker := "?";
END_CASE
q_sDelay := WCONCAT(TO_WSTRING(TIME_TO_UDINT(i_stSet.tLostDelay) / 1000), " s");

q_bWatch := FALSE;
IF _n >= 1 AND _n <= 3 THEN
	q_bWatch := i_abUse[_n];
END_IF
IF q_bWatch THEN
	_tonLost(IN := NOT i_abConnected[_n], PT := i_stSet.tLostDelay);
ELSE
	_tonLost(IN := FALSE);
END_IF
q_bLost := _tonLost.Q;

q_bToManual := q_bLost AND NOT _bDone AND i_bActive;
IF q_bToManual THEN
	_bDone := TRUE;
END_IF
IF NOT q_bLost THEN
	_bDone := FALSE;		// 다시 접속: 다음 끊김에 다시 한 번
END_IF

END_FUNCTION_BLOCK

// ---- 20_Module/Virtual/PRG_SimLink.TcPOU
PROGRAM PRG_SimLink		// 가상 장비끼리 연결 (사무실 시험 전용)
VAR_TEMP
	u			: UINT;
	p			: UINT;
	stUnit		: ST_UnitState;
	fP			: REAL;
	fQ			: REAL;
	b			: UINT;
	afPBat		: ARRAY[1..GVL_PARAM.BAT_COUNT] OF REAL;	// kW, 배터리 그룹(DC 버스)마다 유닛 P 합
END_VAR

(* 실제 현장에서 전기가 이어 주는 것을 흉내 냄: PCS 출력 → 배터리 SOC, 접속점 계측
   - 가상 PCS 여러 대(GVL_SITE.g_aipPcs) → 배터리 그룹마다 그 그룹 BMS (GVL_SITE.BMS_CFG), 계측기1 하나 기준
   - BMS를 늘리거나 줄이면 아래 BMS 줄도 같이 맞춤
   - 현장 빌드: GVL_SITE의 장비를 실제 드라이버로 바꾸고, MAIN의 PRG_SimLink() 호출과 Virtual 폴더 삭제 *)
fP := 0;
fQ := 0;
FOR b := 1 TO GVL_PARAM.BAT_COUNT DO
	afPBat[b] := 0;
END_FOR
FOR u := 1 TO GVL_PARAM.UNIT_COUNT DO
	p := GVL_SITE.UNIT_CFG[u].nPcs;
	IF p >= 1 AND p <= GVL_PARAM.PCS_COUNT THEN
		IF GVL_SITE.g_aipPcs[p] <> 0 THEN
			stUnit	:= GVL_SITE.g_aipPcs[p].M_GetUnitState(GVL_SITE.UNIT_CFG[u].nSub);
			fP		:= fP + stUnit.stP.fValue;
			fQ		:= fQ + stUnit.stQ.fValue;
			b		:= GVL_SITE.UNIT_CFG[u].nBatGroup;
			IF b >= 1 AND b <= GVL_PARAM.BAT_COUNT THEN
				afPBat[b] := afPBat[b] + stUnit.stP.fValue;
			END_IF
		END_IF
	END_IF
END_FOR
// BMS1: physical-map driver has no simulated power input.
// BMS2: physical-map driver has no simulated power input.
// BMS3: physical-map driver has no simulated power input.
GVL_SITE.g_fbMeter1.i_fP	:= fP;
GVL_SITE.g_fbMeter1.i_fQ	:= fQ;

END_PROGRAM

// ---- 99_Test/PRG_TestCtrlMode.TcPOU
PROGRAM PRG_TestCtrlMode		// 제어 모드 자동 시험 (GVL_SITE.TEST_MODE일 때 MAIN이 부름). 실제 제어와 따로 둔 인스턴스만 씀 (장비 지령에 영향 없음)
// 온라인에서 bDone = TRUE가 되면 fbTally.q_nPass·q_nFail, 실패하면 fbTally.q_anFail(실패한 시험 번호)을 봄. bRestart := TRUE로 다시 돌림
// 1~16: 스케줄 모드 단위 시험 (한 스캔). 20~32: 관리자 전환 시험 (여러 스캔, 약 3 s)
VAR
	bRestart	: BOOL;			// TRUE로 쓰면 처음부터 다시
	bDone		: BOOL;			// 시험 끝
	nStep		: UINT;
	fbTally		: FB_TestTally;
	fbSched		: FB_CmSchedule		:= (i_nModuleId := 9001, i_sName := 'TestSched');
	fbConst		: FB_CmConstPower	:= (i_nModuleId := 9002, i_sName := 'TestConst');
	fbMgr		: FB_CtrlModeMgr	:= (i_nModuleId := 9000, i_sName := 'TestMgr');
	aipMode		: ARRAY[1..GVL_PARAM.CTRL_MODE_COUNT] OF I_ControlMode;	// 1 = 정출력 50 kW, 2 = 스케줄
	stCommon	: ST_CmCommonSet;
	stTable		: ST_CmScheduleSet;
	stView		: ST_CtrlModeView;
	stOut		: ST_CtrlModeOut;
	stMgrOut	: ST_SourceOutput;
	stReg		: ST_SourceReg := (bEnable := TRUE, nGrade := 1, ePowerMode := E_SourceMode.Auto, nGroup := 0, tExpire := T#10S);
	tonWait		: TON;
	wsTmp		: WSTRING(63);
END_VAR

IF bRestart THEN
	bRestart	:= FALSE;
	bDone		:= FALSE;
	nStep		:= 0;
END_IF

CASE nStep OF
	0:	// 준비 + 스케줄 단위 시험 (한 스캔)
		fbTally.M_Reset();
		A_Setup();
		A_UnitSchedule();
		fbMgr.i_nModeReq := 2;
		nStep := 10;

	10:	// 관리자: 모드 없음 → 스케줄(2). 켜진 모드가 없으므로 바로 진입
		A_CycleMgr();
		fbTally.M_Check(i_nId := 20, i_bOk := fbMgr.q_nActive = 2 AND fbMgr.q_eStep = E_CtrlModeStep.Active);
		fbTally.M_Check(i_nId := 21, i_bOk := stMgrOut.bPSetActive AND ABS(stMgrOut.fPSet - 200.0) < 0.01);
		fbMgr.i_nModeReq := 1;
		nStep := 11;

	11:	// 정출력(1) 요청 첫 스캔: 이전 모드 끝, 출력 0으로 전환 중
		A_CycleMgr();
		fbTally.M_Check(i_nId := 22, i_bOk := fbMgr.q_eStep = E_CtrlModeStep.Leaving AND fbMgr.q_nActive = 0 AND fbMgr.q_nTarget = 1);
		fbTally.M_Check(i_nId := 23, i_bOk := stMgrOut.bPSetActive AND ABS(stMgrOut.fPSet) < 0.01);
		nStep := 12;

	12:	// tZeroDelay(1 s) 뒤 정출력 진입
		A_CycleMgr();
		tonWait(IN := TRUE, PT := T#3S);
		IF fbMgr.q_eStep = E_CtrlModeStep.Active OR tonWait.Q THEN
			fbTally.M_Check(i_nId := 24, i_bOk := fbMgr.q_nActive = 1 AND ABS(stMgrOut.fPSet - 50.0) < 0.01);
			fbTally.M_Check(i_nId := 25, i_bOk := tonWait.ET >= T#900MS AND NOT tonWait.Q);
			tonWait(IN := FALSE);
			fbMgr.i_nModeReq := 9;
			nStep := 13;
		END_IF

	13:	// 없는 칸(9) → BadSlot, 지금 모드 유지
		A_CycleMgr();
		fbTally.M_Check(i_nId := 26, i_bOk := fbMgr.q_eRefuse = E_CtrlModeRefuse.BadSlot AND fbMgr.q_nActive = 1);
		stView.stTime.bValid	:= FALSE;
		fbMgr.i_nModeReq		:= 2;
		nStep := 14;

	14:	// 시각 무효 → 스케줄 진입 거부 (NotReady, 이유 NO_TIME), 정출력 유지
		A_CycleMgr();
		fbTally.M_Check(i_nId := 27, i_bOk := fbMgr.q_eRefuse = E_CtrlModeRefuse.NotReady AND fbMgr.q_nRefuseReason = GVL_CM_RSN.NO_TIME AND fbMgr.q_nActive = 1);
		fbTally.M_Check(i_nId := 28, i_bOk := ABS(stMgrOut.fPSet - 50.0) < 0.01);
		stView.stTime.bValid	:= TRUE;
		fbMgr.i_bRetry			:= TRUE;		// 같은 요청(2)을 다시
		nStep := 15;

	15:	// 재시도 → 전환 시작
		A_CycleMgr();
		fbTally.M_Check(i_nId := 29, i_bOk := fbMgr.q_eStep = E_CtrlModeStep.Leaving AND fbMgr.q_nTarget = 2 AND NOT fbMgr.i_bRetry);
		nStep := 16;

	16:	// 스케줄 진입
		A_CycleMgr();
		tonWait(IN := TRUE, PT := T#3S);
		IF fbMgr.q_eStep = E_CtrlModeStep.Active OR tonWait.Q THEN
			fbTally.M_Check(i_nId := 30, i_bOk := fbMgr.q_nActive = 2 AND ABS(stMgrOut.fPSet - 200.0) < 0.01);
			tonWait(IN := FALSE);
			fbMgr.i_nModeReq := 0;
			nStep := 17;
		END_IF

	17:	// 모드 없음(0) → 출력 0 뒤 지령 없음
		A_CycleMgr();
		tonWait(IN := TRUE, PT := T#3S);
		IF fbMgr.q_eStep = E_CtrlModeStep.Idle OR tonWait.Q THEN
			fbTally.M_Check(i_nId := 31, i_bOk := fbMgr.q_eStep = E_CtrlModeStep.Idle AND fbMgr.q_nActive = 0 AND NOT stMgrOut.bPSetActive);
			tonWait(IN := FALSE);
			// 설정 점검: 시작 > 끝인 칸이 있으면 관리자가 모드의 오류 문구를 올림
			stTable.astSlot[2, 3, 5].nStart	:= 1500;
			stTable.astSlot[2, 3, 5].nEnd	:= 1400;
			fbSched.i_stTable := stTable;
			wsTmp := fbMgr.M_CheckSet();
			fbTally.M_Check(i_nId := 32, i_bOk := wsTmp <> "");
			stTable.astSlot[2, 3, 5].nStart	:= 0;
			stTable.astSlot[2, 3, 5].nEnd	:= 0;
			fbSched.i_stTable := stTable;
			wsTmp := fbMgr.M_CheckSet();
			fbTally.M_Check(i_nId := 33, i_bOk := wsTmp = "");
			nStep := 99;
		END_IF

	99:
		bDone := TRUE;
END_CASE

ACTION A_Setup:
// 모드 등록·설정
aipMode[1]	:= fbConst;
aipMode[2]	:= fbSched;
fbConst.i_stSet.fPSet	:= 50.0;
fbConst.i_stSet.bQSet	:= FALSE;
fbConst.i_stSet.tDuration	:= T#0S;
// 공통 설정: 기본값(방전 08:00~22:00, 일요일 금지, 역송 여유 10 kW·0.95) + 7월 14일 휴일
stCommon.abHoliday[7, 14]	:= TRUE;
// 시간표: 여름(0) 월요일(1), 일요일(0)
stTable.astSlot[0, 1, 1].nStart := 100;		stTable.astSlot[0, 1, 1].nEnd := 600;		stTable.astSlot[0, 1, 1].fP := -300.0;	// 충전
stTable.astSlot[0, 1, 2].nStart := 1000;	stTable.astSlot[0, 1, 2].nEnd := 1200;		stTable.astSlot[0, 1, 2].fP := 200.0;	// 방전
stTable.astSlot[0, 1, 3].nStart := 1100;	stTable.astSlot[0, 1, 3].nEnd := 1130;		stTable.astSlot[0, 1, 3].fP := 400.0;	// 겹침: 번호 큰 칸
stTable.astSlot[0, 1, 4].nStart := 2300;	stTable.astSlot[0, 1, 4].nEnd := 2400;		stTable.astSlot[0, 1, 4].fP := 100.0;	// 방전 허용 시간 밖
stTable.astSlot[0, 0, 1].nStart := 1000;	stTable.astSlot[0, 0, 1].nEnd := 1200;		stTable.astSlot[0, 0, 1].fP := 200.0;	// 일요일
fbSched.i_stCommon	:= stCommon;
fbSched.i_stTable	:= stTable;
// 관리자: 기본 설정 (전환 때 1 s 출력 0, 대체 모드 없음)
fbMgr.i_stSet.bZeroOnSwitch	:= TRUE;
fbMgr.i_stSet.tZeroDelay	:= T#1S;
fbMgr.i_stSet.nFallback		:= 0;
fbMgr.i_bRetry				:= FALSE;
A_ViewBase();
END_ACTION

ACTION A_ViewBase:
// 기준 상황: 2026-07-13 월요일 10:30:00, 가용 유닛 1, 가용 출력 1000 kW, 수전 1000 kW (접속점 P = -1000), ESS 출력 0
stView.stTime.bValid		:= TRUE;
stView.stTime.nYear			:= 2026;
stView.stTime.nMonth		:= 7;
stView.stTime.nDay			:= 13;
stView.stTime.nDayOfWeek	:= 1;
stView.stTime.nHour			:= 10;
stView.stTime.nMinute		:= 30;
stView.stTime.nSecond		:= 0;
stView.stGroup.nUnitAvail	:= 1;
stView.stGroup.fPRatedAvail	:= 1000.0;
stView.stGroup.fPOut		:= 0.0;
stView.stGroup.stPcc.stMeas.stP.bValid	:= TRUE;
stView.stGroup.stPcc.stMeas.stP.fValue	:= -1000.0;
END_ACTION

ACTION A_UnitSchedule:
fbSched.M_Enter(i_stView := stView);

// 1) 03:00 충전 칸 → -300
A_ViewBase();
stView.stTime.nHour := 3;	stView.stTime.nMinute := 0;
stOut := fbSched.M_Calc(i_stView := stView);
fbTally.M_Check(i_nId := 1, i_bOk := ABS(stOut.fPSet + 300.0) < 0.01 AND fbSched.q_nSlot = 1 AND fbSched.q_nState = 0);

// 2) 10:30 방전 칸 → 200
A_ViewBase();
stOut := fbSched.M_Calc(i_stView := stView);
fbTally.M_Check(i_nId := 2, i_bOk := ABS(stOut.fPSet - 200.0) < 0.01 AND fbSched.q_nSlot = 2 AND fbSched.q_nState = 0);

// 3) 11:15 겹친 칸 → 번호 큰 칸 400
A_ViewBase();
stView.stTime.nHour := 11;	stView.stTime.nMinute := 15;
stOut := fbSched.M_Calc(i_stView := stView);
fbTally.M_Check(i_nId := 3, i_bOk := ABS(stOut.fPSet - 400.0) < 0.01 AND fbSched.q_nSlot = 3);

// 4) 12:00 = 끝 시각 (미포함) → 칸 없음 0, 지령은 냄
A_ViewBase();
stView.stTime.nHour := 12;	stView.stTime.nMinute := 0;
stOut := fbSched.M_Calc(i_stView := stView);
fbTally.M_Check(i_nId := 4, i_bOk := stOut.bPSetActive AND ABS(stOut.fPSet) < 0.01 AND fbSched.q_nSlot = 0 AND fbSched.q_nState = GVL_CM_RSN.NO_SLOT);

// 5) 23:30 방전 칸이지만 방전 허용 시간 밖 → 0
A_ViewBase();
stView.stTime.nHour := 23;
stOut := fbSched.M_Calc(i_stView := stView);
fbTally.M_Check(i_nId := 5, i_bOk := ABS(stOut.fPSet) < 0.01 AND fbSched.q_nSlot = 4 AND fbSched.q_nState = GVL_CM_RSN.DIS_TIME);

// 6) 일요일 10:30 방전 칸 → 일요일 방전 금지로 0
A_ViewBase();
stView.stTime.nDayOfWeek := 0;	stView.stTime.nDay := 12;
stOut := fbSched.M_Calc(i_stView := stView);
fbTally.M_Check(i_nId := 6, i_bOk := ABS(stOut.fPSet) < 0.01 AND fbSched.q_nSlot = 1 AND fbSched.q_nState = GVL_CM_RSN.DIS_TIME);

// 7) 역송 방지: 수전 150 kW → 부하 150, 가능 140 → 140 × 0.95 = 133
A_ViewBase();
stView.stGroup.stPcc.stMeas.stP.fValue := -150.0;
stOut := fbSched.M_Calc(i_stView := stView);
fbTally.M_Check(i_nId := 7, i_bOk := ABS(stOut.fPSet - 133.0) < 0.01 AND fbSched.q_nState = GVL_CM_RSN.REV_LIMIT);

// 8) 접속점 계측 무효 → 방전 0
A_ViewBase();
stView.stGroup.stPcc.stMeas.stP.bValid := FALSE;
stOut := fbSched.M_Calc(i_stView := stView);
fbTally.M_Check(i_nId := 8, i_bOk := ABS(stOut.fPSet) < 0.01 AND fbSched.q_nState = GVL_CM_RSN.NO_PCC);

// 9) 휴일 (7월 14일) → 0
A_ViewBase();
stView.stTime.nDay := 14;	stView.stTime.nDayOfWeek := 2;
stOut := fbSched.M_Calc(i_stView := stView);
fbTally.M_Check(i_nId := 9, i_bOk := ABS(stOut.fPSet) < 0.01 AND fbSched.q_nState = GVL_CM_RSN.HOLIDAY);

// 10) 시각 무효 → 0, 진입 거부 이유 NO_TIME
A_ViewBase();
stView.stTime.bValid := FALSE;
stOut := fbSched.M_Calc(i_stView := stView);
fbTally.M_Check(i_nId := 10, i_bOk := ABS(stOut.fPSet) < 0.01 AND fbSched.q_nState = GVL_CM_RSN.NO_TIME AND fbSched.M_CheckEnter(i_stView := stView) = GVL_CM_RSN.NO_TIME);

// 11) 1월 = 겨울(2): 겨울 시간표가 비어 칸 없음
A_ViewBase();
stView.stTime.nMonth := 1;
stOut := fbSched.M_Calc(i_stView := stView);
fbTally.M_Check(i_nId := 11, i_bOk := fbSched.q_nSeason = 2 AND fbSched.q_nState = GVL_CM_RSN.NO_SLOT);

// 12) ESS 충전 중 역송 방지: 수전 500, ESS -300 → 부하 200, 가능 190 → 180.5
A_ViewBase();
stView.stGroup.stPcc.stMeas.stP.fValue := -500.0;
stView.stGroup.fPOut := -300.0;
stOut := fbSched.M_Calc(i_stView := stView);
fbTally.M_Check(i_nId := 12, i_bOk := ABS(stOut.fPSet - 180.5) < 0.01 AND fbSched.q_nState = GVL_CM_RSN.REV_LIMIT);

// 13) 진입 검사: 정상이면 0
A_ViewBase();
fbTally.M_Check(i_nId := 13, i_bOk := fbSched.M_CheckEnter(i_stView := stView) = 0);

// 14) 설정 점검: 시작 > 끝인 칸 → 오류 문구, 되돌리면 정상
stTable.astSlot[1, 4, 2].nStart := 1300;	stTable.astSlot[1, 4, 2].nEnd := 1200;
fbSched.i_stTable := stTable;
wsTmp := fbSched.M_CheckSet();
fbTally.M_Check(i_nId := 14, i_bOk := wsTmp <> "");
stTable.astSlot[1, 4, 2].nStart := 0;		stTable.astSlot[1, 4, 2].nEnd := 0;
fbSched.i_stTable := stTable;
wsTmp := fbSched.M_CheckSet();
fbTally.M_Check(i_nId := 15, i_bOk := wsTmp = "");

// 16) 방전 허용 시간을 끄면 23:30 방전 칸 100
stCommon.stDis.bUse := FALSE;
fbSched.i_stCommon := stCommon;
A_ViewBase();
stView.stTime.nHour := 23;
stOut := fbSched.M_Calc(i_stView := stView);
fbTally.M_Check(i_nId := 16, i_bOk := ABS(stOut.fPSet - 100.0) < 0.01 AND fbSched.q_nState = 0);
stCommon.stDis.bUse := TRUE;
fbSched.i_stCommon := stCommon;

// 17) 진입 검사: 가용 유닛 없음 → NO_UNIT
A_ViewBase();
stView.stGroup.nUnitAvail := 0;
fbTally.M_Check(i_nId := 17, i_bOk := fbSched.M_CheckEnter(i_stView := stView) = GVL_CM_RSN.NO_UNIT);

fbSched.M_Exit();
A_ViewBase();
END_ACTION

ACTION A_CycleMgr:
// 관리자 한 스캔 (FB_SourceHub가 하는 것처럼 M_Cycle을 부름)
fbMgr.i_aipMode	:= aipMode;
fbMgr.i_stTime	:= stView.stTime;
fbMgr.M_Cycle(i_stReg := stReg, i_stView := stView.stGroup);
stMgrOut := fbMgr.Output;
END_ACTION

END_PROGRAM

// ---- 99_Test/FB_TestTally.TcPOU
FUNCTION_BLOCK FB_TestTally		// 시험 결과 세기: 통과·실패 수와 실패한 시험 번호
VAR_OUTPUT
	q_nPass		: UINT;
	q_nFail		: UINT;
	q_anFail	: ARRAY[1..32] OF UINT;		// 실패한 시험 번호 (앞에서부터)
END_VAR

METHOD M_Reset
VAR
	nI	: UINT;
END_VAR
q_nPass := 0;
q_nFail := 0;
FOR nI := 1 TO 32 DO
	q_anFail[nI] := 0;
END_FOR
END_METHOD

METHOD M_Check : BOOL
VAR_INPUT
	i_nId	: UINT;		// 시험 번호
	i_bOk	: BOOL;
END_VAR
IF i_bOk THEN
	q_nPass := q_nPass + 1;
ELSE
	q_nFail := q_nFail + 1;
	IF q_nFail <= 32 THEN
		q_anFail[q_nFail] := i_nId;
	END_IF
END_IF
M_Check := i_bOk;
END_METHOD

END_FUNCTION_BLOCK

// ---- 20_Module/ControlMode/FB_CmSchedule.TcPOU
FUNCTION_BLOCK FB_CmSchedule EXTENDS FB_CmTariffBase		// 제어 모드: 스케줄 (Messis SCHEDULE_MODE). 계절·요일 시간표의 P를 냄
// 맞는 칸 없음·휴일·시각 무효 → 0. 충전(-)은 그대로, 방전(+)은 방전 허용 시간·역송 방지 (공통 설정). 칸은 자정을 넘지 않음
VAR_INPUT
	i_stTable	: ST_CmScheduleSet;		// 시간표 (A_PassModuleSet이 GVL_PERSIST.g_stModuleSet.stCmSchedule을 매 스캔 넘김)
END_VAR

METHOD M_Calc : ST_CtrlModeOut
VAR_INPUT
	i_stView	: ST_CtrlModeView;
END_VAR
VAR
	fP		: REAL;
	nRsn	: UINT;
END_VAR
fP := 0.0;
IF M_Begin(i_stView := i_stView) THEN
	M_SchedLookup(i_stTime := i_stView.stTime, iq_stTable := i_stTable);
	fP			:= M_SchedOut(i_stView := i_stView, q_nRsn => nRsn);
	q_nState	:= nRsn;
END_IF
M_Calc := M_Finish(i_fP := fP);
END_METHOD

METHOD M_CheckSet : WSTRING(63)
M_CheckSet := SUPER^.M_CheckSet();
IF M_CheckSet = "" THEN
	M_CheckSet := M_CheckTable(iq_stTable := i_stTable);
END_IF
END_METHOD

END_FUNCTION_BLOCK

// ---- 20_Module/ControlMode/FB_CmTariffBase.TcPOU
FUNCTION_BLOCK ABSTRACT FB_CmTariffBase EXTENDS FB_CtrlModeBase		// 요금제 기반 제어 모드 공통 바탕 (스케줄·피크컷·통합). 같은 계산은 여기 메서드 하나만 씀
// 휴일·계절·방전 허용 시간·역송 방지·시간표 조회·잔량 방전·자동 충전. 상태·이유 코드는 GVL_CM_RSN
// 파생 FB: M_Calc에서 M_Begin으로 시작 → 계산 → M_Finish로 끝냄
VAR_INPUT
	i_stCommon	: ST_CmCommonSet;	// 공통 설정 (A_PassModuleSet이 GVL_PERSIST.g_stModuleSet.stCmCommon을 매 스캔 넘김)
END_VAR
VAR_OUTPUT
	q_nState	: UINT;		// 0 = 정상, 그 외 = GVL_CM_RSN (M_ReasonText)
	q_fOutP		: REAL;		// 이번 스캔에 낸 P (kW, 방전 +)
	q_nSeason	: UINT;		// 지금 계절 (0 여름, 1 봄·가을, 2 겨울)
	q_nSlot		: UINT;		// 맞는 시간표 칸 (0 = 없음, 시간표를 쓰는 모드만)
	q_fSlotP	: REAL;		// 그 칸 값 (kW)
END_VAR

METHOD M_CheckEnter : UINT
VAR_INPUT
	i_stView	: ST_CtrlModeView;
END_VAR
M_CheckEnter := 0;
IF NOT M_TimeOk(i_stTime := i_stView.stTime) THEN
	M_CheckEnter := GVL_CM_RSN.NO_TIME;
ELSIF i_stView.stGroup.nUnitAvail = 0 THEN
	M_CheckEnter := GVL_CM_RSN.NO_UNIT;
END_IF
END_METHOD

METHOD PROTECTED M_Begin : BOOL		// 스캔 시작: 출력 칸을 비우고 계절을 셈. 시각이 맞고 휴일이 아니면 TRUE (FALSE면 q_nState에 이유, 0을 냄)
VAR_INPUT
	i_stView	: ST_CtrlModeView;
END_VAR
q_nState	:= 0;
q_fOutP		:= 0.0;
q_nSlot		:= 0;
q_fSlotP	:= 0.0;
M_Begin		:= FALSE;
IF NOT M_TimeOk(i_stTime := i_stView.stTime) THEN
	q_nState := GVL_CM_RSN.NO_TIME;
ELSE
	q_nSeason := i_stCommon.anSeasonOfMonth[i_stView.stTime.nMonth];
	IF q_nSeason > 2 THEN
		q_nSeason := 0;		// M_CheckSet이 막지만 배열 범위 보호
	END_IF
	IF i_stCommon.abHoliday[i_stView.stTime.nMonth, i_stView.stTime.nDay] THEN
		q_nState := GVL_CM_RSN.HOLIDAY;
	ELSE
		M_Begin := TRUE;
	END_IF
END_IF
END_METHOD

METHOD PROTECTED M_Finish : ST_CtrlModeOut		// 스캔 끝: P를 지령으로 냄 (0이어도 냄: 등급이 낮은 지령원으로 넘어가지 않게). Q는 내지 않음
VAR_INPUT
	i_fP		: REAL;		// kW, 방전 +
END_VAR
q_fOutP					:= i_fP;
M_Finish.bPSetActive	:= TRUE;
M_Finish.fPSet			:= i_fP;
M_Finish.bQSetActive	:= FALSE;
M_Finish.fQSet			:= 0.0;
M_Finish.bExitReq		:= FALSE;
M_Finish.nReason		:= 0;
END_METHOD

METHOD PROTECTED M_TimeOk : BOOL		// 시각이 유효하고 배열 번호로 쓸 수 있는 범위
VAR_INPUT
	i_stTime	: ST_LocalTime;
END_VAR
M_TimeOk := i_stTime.bValid AND i_stTime.nMonth >= 1 AND i_stTime.nMonth <= 12
	AND i_stTime.nDay >= 1 AND i_stTime.nDay <= 31 AND i_stTime.nDayOfWeek <= 6;
END_METHOD

METHOD PROTECTED M_DisAllowed : BOOL		// 지금 방전해도 되는 시간인가 (공통 설정 stDis)
VAR_INPUT
	i_stTime	: ST_LocalTime;
END_VAR
M_DisAllowed := TRUE;
IF i_stCommon.stDis.bUse THEN
	M_DisAllowed := F_InHhmmWindow(i_nNow := F_TimeHhmm(i_stTime := i_stTime), i_nStart := i_stCommon.stDis.nStart, i_nEnd := i_stCommon.stDis.nEnd)
		AND (i_stTime.nDayOfWeek <> 0 OR i_stCommon.stDis.bSunday);
END_IF
END_METHOD

METHOD PROTECTED M_NoReverse : REAL		// 역송 방지: 방전 요청을 (부하 − 여유) 안으로 줄임 (공통 설정 stNoRev). 충전·0은 그대로
VAR_INPUT
	i_fReq		: REAL;		// kW, 방전 +
	i_stView	: ST_CtrlModeView;
END_VAR
VAR_OUTPUT
	q_nRsn		: UINT;		// 0 = 그대로, GVL_CM_RSN.REV_LIMIT = 줄임, GVL_CM_RSN.NO_PCC = 계측 무효로 0
END_VAR
VAR
	fLoad		: REAL;		// 부하 = ESS가 없을 때의 수전
	fAvail		: REAL;		// 역송 없이 방전할 수 있는 양
END_VAR
M_NoReverse	:= i_fReq;
q_nRsn		:= 0;
IF i_fReq > 0.0 AND i_stCommon.stNoRev.bUse THEN
	IF i_stView.stGroup.stPcc.stMeas.stP.bValid THEN
		// 접속점 P는 공급(역송) +, 수전 -. 부하 = ESS 출력 − 접속점 공급 (충전 중·역송 중에도 맞음)
		fLoad	:= MAX(i_stView.stGroup.fPOut - i_stView.stGroup.stPcc.stMeas.stP.fValue, 0.0);
		fAvail	:= MAX(fLoad - i_stCommon.stNoRev.fMargin, 0.0);
		IF i_fReq > fAvail THEN
			M_NoReverse	:= fAvail * i_stCommon.stNoRev.fScale;
			q_nRsn		:= GVL_CM_RSN.REV_LIMIT;
		END_IF
	ELSE
		M_NoReverse	:= 0.0;
		q_nRsn		:= GVL_CM_RSN.NO_PCC;
	END_IF
END_IF
END_METHOD

METHOD PROTECTED M_SchedLookup : BOOL		// 시간표에서 지금 맞는 칸 (번호가 큰 칸 우선). 찾으면 TRUE, q_nSlot·q_fSlotP에 씀. M_Begin 뒤에 부름 (계절)
VAR_INPUT
	i_stTime	: ST_LocalTime;
END_VAR
VAR_IN_OUT CONSTANT
	iq_stTable	: ST_CmScheduleSet;
END_VAR
VAR
	nNow		: UINT;
	k			: UINT;
END_VAR
nNow		:= F_TimeHhmm(i_stTime := i_stTime);
q_nSlot		:= 0;
q_fSlotP	:= 0.0;
FOR k := 1 TO GVL_PARAM.SCHED_SLOT_COUNT DO
	IF F_InHhmmWindow(i_nNow := nNow, i_nStart := iq_stTable.astSlot[q_nSeason, i_stTime.nDayOfWeek, k].nStart, i_nEnd := iq_stTable.astSlot[q_nSeason, i_stTime.nDayOfWeek, k].nEnd) THEN
		q_nSlot		:= k;
		q_fSlotP	:= iq_stTable.astSlot[q_nSeason, i_stTime.nDayOfWeek, k].fP;
	END_IF
END_FOR
M_SchedLookup := q_nSlot <> 0;
END_METHOD

METHOD PROTECTED M_SchedOut : REAL		// 시간표 값 → 낼 값: 칸 없음 0, 충전 그대로, 방전은 방전 허용 시간·역송 방지 (스케줄·통합 모드 공통)
VAR_INPUT
	i_stView	: ST_CtrlModeView;
END_VAR
VAR_OUTPUT
	q_nRsn		: UINT;		// 0 = 칸 값 그대로, 그 외 GVL_CM_RSN
END_VAR
q_nRsn		:= 0;
M_SchedOut	:= 0.0;
IF q_nSlot = 0 THEN
	q_nRsn := GVL_CM_RSN.NO_SLOT;
ELSIF q_fSlotP > 0.0 THEN
	IF M_DisAllowed(i_stTime := i_stView.stTime) THEN
		M_SchedOut := M_NoReverse(i_fReq := q_fSlotP, i_stView := i_stView, q_nRsn => q_nRsn);
	ELSE
		q_nRsn := GVL_CM_RSN.DIS_TIME;
	END_IF
ELSE
	M_SchedOut := q_fSlotP;		// 충전 (또는 0)
END_IF
END_METHOD

METHOD PROTECTED M_RemainDis : REAL		// 잔량 방전량 (kW): (지금 에너지 − 하한 SOC 에너지)를 끝 시각까지 고르게. 가용 출력 상한. 역송 방지 전
VAR_INPUT
	i_stView	: ST_CtrlModeView;
	i_stWin		: ST_CmWindowSet;	// nEnd, fSoc = 남길 하한
END_VAR
VAR_OUTPUT
	q_bNoCap	: BOOL;		// 용량·SOC 무효
END_VAR
VAR
	nMin		: UINT;
	fE			: REAL;		// kWh
END_VAR
M_RemainDis	:= 0.0;
q_bNoCap	:= i_stView.stGroup.fCapacity <= 0.0 OR NOT i_stView.stGroup.stSocAvg.bValid;
IF NOT q_bNoCap THEN
	nMin	:= F_MinutesTo(i_nNow := F_TimeHhmm(i_stTime := i_stView.stTime), i_nEnd := i_stWin.nEnd);
	fE		:= i_stView.stGroup.fCapacity * (i_stView.stGroup.stSocAvg.fValue - i_stWin.fSoc) / 100.0;
	IF nMin > 0 AND fE > 0.0 THEN
		M_RemainDis := MIN(fE * 60.0 / UINT_TO_REAL(nMin), i_stView.stGroup.fPRatedAvail);
	END_IF
END_IF
END_METHOD

METHOD PROTECTED M_AutoChg : REAL		// 자동 충전량 (kW, 양수): (목표 SOC 에너지 − 지금 에너지)를 끝 시각까지 + 1 kW, 최소 10 kW, 가용 출력 상한
VAR_INPUT
	i_stView	: ST_CtrlModeView;
	i_stWin		: ST_CmWindowSet;	// nEnd, fSoc = 채울 목표
END_VAR
VAR_OUTPUT
	q_bNoCap	: BOOL;		// 용량·SOC 무효
END_VAR
VAR
	nMin		: UINT;
	fE			: REAL;		// kWh
END_VAR
M_AutoChg	:= 0.0;
q_bNoCap	:= i_stView.stGroup.fCapacity <= 0.0 OR NOT i_stView.stGroup.stSocAvg.bValid;
IF NOT q_bNoCap THEN
	nMin	:= F_MinutesTo(i_nNow := F_TimeHhmm(i_stTime := i_stView.stTime), i_nEnd := i_stWin.nEnd);
	fE		:= i_stView.stGroup.fCapacity * (i_stWin.fSoc - i_stView.stGroup.stSocAvg.fValue) / 100.0;
	IF nMin > 0 AND fE > 0.0 THEN
		M_AutoChg := MIN(MAX(fE * 60.0 / UINT_TO_REAL(nMin) + 1.0, 10.0), i_stView.stGroup.fPRatedAvail);
	END_IF
END_IF
END_METHOD

METHOD PROTECTED M_CheckTable : WSTRING(63)		// 시간표 칸 시각 점검 (시작 ≤ 끝, HHMM)
VAR_IN_OUT CONSTANT
	iq_stTable	: ST_CmScheduleSet;
END_VAR
VAR
	nS	: UINT;		// 계절
	nD	: UINT;		// 요일
	nK	: UINT;		// 칸
END_VAR
M_CheckTable := "";
FOR nS := 0 TO 2 DO
	FOR nD := 0 TO 6 DO
		FOR nK := 1 TO GVL_PARAM.SCHED_SLOT_COUNT DO
			IF NOT F_RealOk(iq_stTable.astSlot[nS, nD, nK].fP) THEN	// [결함 13 수정 2026-11-04: 칸 출력 kW가 숫자가 아님]
				M_CheckTable := WCONCAT(WCONCAT(WCONCAT(WCONCAT(WCONCAT("시간표 칸 출력 숫자 아님: 계절 ", TO_WSTRING(nS)), " 요일 "), TO_WSTRING(nD)), " 칸 "), TO_WSTRING(nK));
				RETURN;
			END_IF
			IF NOT F_HhmmOk(i_nHhmm := iq_stTable.astSlot[nS, nD, nK].nStart) OR NOT F_HhmmOk(i_nHhmm := iq_stTable.astSlot[nS, nD, nK].nEnd)
				OR iq_stTable.astSlot[nS, nD, nK].nStart > iq_stTable.astSlot[nS, nD, nK].nEnd THEN
				M_CheckTable := WCONCAT(WCONCAT(WCONCAT(WCONCAT(WCONCAT("시간표 칸 시각 잘못됨: 계절 ", TO_WSTRING(nS)), " 요일 "), TO_WSTRING(nD)), " 칸 "), TO_WSTRING(nK));
				RETURN;
			END_IF
		END_FOR
	END_FOR
END_FOR
END_METHOD

METHOD PROTECTED M_CheckWindow : BOOL		// 시간 구간 설정이 맞는가 (쓰지 않으면 TRUE)
VAR_INPUT
	i_stWin		: ST_CmWindowSet;
END_VAR
// [결함 13 수정 2026-11-04: SOC가 숫자가 아니면 (쓰지 않는 구간이어도) 틀림. 비교 전에 비트로. 원래 NOT i_stWin.bUse OR (… AND i_stWin.fSoc >= 0.0 AND i_stWin.fSoc <= 100.0)]
IF NOT F_RealOk(i_stWin.fSoc) THEN
	M_CheckWindow := FALSE;
	RETURN;
END_IF
M_CheckWindow := NOT i_stWin.bUse OR (F_HhmmOk(i_nHhmm := i_stWin.nStart) AND F_HhmmOk(i_nHhmm := i_stWin.nEnd)
	AND i_stWin.nStart <> i_stWin.nEnd AND i_stWin.fSoc >= 0.0 AND i_stWin.fSoc <= 100.0);
END_METHOD

METHOD M_ReasonText : WSTRING(63)
VAR_INPUT
	i_nReason	: UINT;
END_VAR
CASE i_nReason OF
	GVL_CM_RSN.NO_TIME:		M_ReasonText := "시각 무효";
	GVL_CM_RSN.NO_UNIT:		M_ReasonText := "가용 유닛 없음";
	GVL_CM_RSN.HOLIDAY:		M_ReasonText := "휴일";
	GVL_CM_RSN.NO_SLOT:		M_ReasonText := "맞는 시간표 칸 없음";
	GVL_CM_RSN.DIS_TIME:	M_ReasonText := "방전 허용 시간 아님";
	GVL_CM_RSN.REV_LIMIT:	M_ReasonText := "역송 방지로 방전 줄임";
	GVL_CM_RSN.NO_PCC:		M_ReasonText := "접속점 계측 무효 (방전 0)";
	GVL_CM_RSN.NO_CAP:		M_ReasonText := "배터리 용량·SOC 무효";
	GVL_CM_RSN.PEAK:		M_ReasonText := "피크 제어 방전";
	GVL_CM_RSN.BELOW_PEAK:	M_ReasonText := "피크 제어 필요 없음";
	GVL_CM_RSN.AUTO_CHG:	M_ReasonText := "자동 충전 시간";
	GVL_CM_RSN.REMAIN_DIS:	M_ReasonText := "잔량 방전 시간";
	GVL_CM_RSN.SCHED_PEAK:	M_ReasonText := "스케줄·피크 제어 중 큰 방전";
	GVL_CM_RSN.NEW_INTERVAL:	M_ReasonText := "새 15분 구간 시작";
ELSE
	M_ReasonText := WCONCAT("이유 ", TO_WSTRING(i_nReason));
END_CASE
END_METHOD

METHOD M_CheckSet : WSTRING(63)		// 공통 설정 점검. 파생 FB는 SUPER^.M_CheckSet() 뒤에 자기 설정을 점검
VAR
	k	: UINT;
END_VAR
M_CheckSet := "";
FOR k := 1 TO 12 DO
	IF i_stCommon.anSeasonOfMonth[k] > 2 THEN
		M_CheckSet := "제어 모드 공통: 월 → 계절 값은 0~2";
		RETURN;
	END_IF
END_FOR
IF NOT F_HhmmOk(i_nHhmm := i_stCommon.stDis.nStart) OR NOT F_HhmmOk(i_nHhmm := i_stCommon.stDis.nEnd) THEN
	M_CheckSet := "제어 모드 공통: 방전 허용 시간 HHMM";
ELSIF NOT (F_RealOk(i_stCommon.stNoRev.fMargin) AND F_RealOk(i_stCommon.stNoRev.fScale)) THEN	// [결함 13 수정 2026-11-04]
	M_CheckSet := "제어 모드 공통: 역송 방지 값 숫자 아님";
ELSIF i_stCommon.stNoRev.fMargin < 0.0 OR i_stCommon.stNoRev.fScale < 0.0 OR i_stCommon.stNoRev.fScale > 1.0 THEN
	M_CheckSet := "제어 모드 공통: 역송 방지 여유 0 이상, 비율 0~1";
END_IF
END_METHOD

END_FUNCTION_BLOCK

// ---- 10_Core/03_Base/FB_CtrlModeBase.TcPOU
FUNCTION_BLOCK ABSTRACT FB_CtrlModeBase EXTENDS FB_ModuleBase IMPLEMENTS I_ControlMode	// 제어 모드 공통 바탕. 파생 FB는 M_Calc만 쓰면 됨 (필요하면 M_CheckEnter·M_Enter·M_Exit·M_ReasonText·M_CheckSet을 바꿈)
// M_Enter·M_Exit를 바꾸면 SUPER^.M_Enter(i_stView := i_stView)·SUPER^.M_Exit()도 부름 (_bActive 유지)
VAR
	_bActive	: BOOL;		// 켜져 있음 (M_Enter ~ M_Exit). 진단용
END_VAR

METHOD M_CheckEnter : UINT		// 기본: 조건 없음
VAR_INPUT
	i_stView	: ST_CtrlModeView;	// 그룹 값(stGroup)·현지 시각(stTime). 관리자가 매 스캔 채움
END_VAR
M_CheckEnter := 0;
END_METHOD

METHOD M_Enter
VAR_INPUT
	i_stView	: ST_CtrlModeView;	// 그룹 값(stGroup)·현지 시각(stTime). 관리자가 매 스캔 채움
END_VAR
_bActive := TRUE;
END_METHOD

METHOD ABSTRACT M_Calc : ST_CtrlModeOut
VAR_INPUT
	i_stView	: ST_CtrlModeView;	// 그룹 값(stGroup)·현지 시각(stTime). 관리자가 매 스캔 채움
END_VAR
END_METHOD

METHOD M_Exit
_bActive := FALSE;
END_METHOD

END_FUNCTION_BLOCK

// ---- 10_Core/02_Util/F_InHhmmWindow.TcPOU
FUNCTION F_InHhmmWindow : BOOL		// 지금이 시간 구간 안인가: 시작 ≤ 지금 < 끝 (HHMM). 시작 > 끝이면 자정을 넘는 구간, 시작 = 끝이면 빈 구간
VAR_INPUT
	i_nNow		: UINT;		// HHMM
	i_nStart	: UINT;
	i_nEnd		: UINT;
END_VAR

IF i_nStart = i_nEnd THEN
	F_InHhmmWindow := FALSE;
ELSIF i_nStart < i_nEnd THEN
	F_InHhmmWindow := i_nNow >= i_nStart AND i_nNow < i_nEnd;
ELSE
	F_InHhmmWindow := i_nNow >= i_nStart OR i_nNow < i_nEnd;
END_IF

END_FUNCTION

// ---- 10_Core/02_Util/F_TimeHhmm.TcPOU
FUNCTION F_TimeHhmm : UINT		// 현지 시각 → HHMM (예: 13시 5분 = 1305)
VAR_INPUT
	i_stTime	: ST_LocalTime;
END_VAR

F_TimeHhmm := i_stTime.nHour * 100 + i_stTime.nMinute;

END_FUNCTION

// ---- 10_Core/02_Util/F_MinutesTo.TcPOU
FUNCTION F_MinutesTo : UINT		// 지금(HHMM)부터 끝(HHMM)까지 남은 분. 끝이 지났으면 다음 날 그 시각까지 (자정을 넘김). 같으면 0
VAR_INPUT
	i_nNow		: UINT;		// HHMM
	i_nEnd		: UINT;		// HHMM (2400 = 자정)
END_VAR
VAR
	nDiff		: DINT;
END_VAR

nDiff := (UINT_TO_DINT(i_nEnd / 100) * 60 + UINT_TO_DINT(i_nEnd MOD 100)) - (UINT_TO_DINT(i_nNow / 100) * 60 + UINT_TO_DINT(i_nNow MOD 100));
IF nDiff < 0 THEN
	nDiff := nDiff + 1440;
END_IF
F_MinutesTo := DINT_TO_UINT(nDiff);

END_FUNCTION

// ---- 10_Core/02_Util/F_HhmmOk.TcPOU
FUNCTION F_HhmmOk : BOOL		// HHMM 값이 맞는가: 0000~2359, 또는 2400 (하루 끝)
VAR_INPUT
	i_nHhmm		: UINT;
END_VAR

F_HhmmOk := ((i_nHhmm / 100) < 24 AND (i_nHhmm MOD 100) < 60) OR i_nHhmm = 2400;

END_FUNCTION

// ---- 20_Module/ControlMode/FB_CmConstPower.TcPOU
FUNCTION_BLOCK FB_CmConstPower EXTENDS FB_CtrlModeBase		// 제어 모드 예: 정출력. 설정한 P(·Q)를 접속점 기준으로 냄. tDuration이 지나면 스스로 끝냄
// 새 제어 모드의 본보기: FB_CtrlModeBase 상속 → M_Calc (+ 필요하면 M_CheckEnter·M_Enter·M_Exit·M_ReasonText·M_CheckSet)
VAR_INPUT
	i_stSet		: ST_CmConstPowerSet;	// 설정 (A_PassModuleSet이 GVL_PERSIST.g_stModuleSet 칸을 매 스캔 넘김)
END_VAR
VAR
	_tonRun		: TON;		// 운전 시간
END_VAR
VAR CONSTANT
	RSN_NO_UNIT	: UINT := 1;	// 진입 거부: 가용 유닛 없음
	RSN_TIME_UP	: UINT := 2;	// 끝: 운전 시간 끝
END_VAR

METHOD M_CheckEnter : UINT
VAR_INPUT
	i_stView	: ST_CtrlModeView;	// 그룹 값(stGroup)·현지 시각(stTime). 관리자가 매 스캔 채움
END_VAR
M_CheckEnter := 0;
IF i_stView.stGroup.nUnitAvail = 0 THEN
	M_CheckEnter := RSN_NO_UNIT;
END_IF
END_METHOD

METHOD M_Enter
VAR_INPUT
	i_stView	: ST_CtrlModeView;	// 그룹 값(stGroup)·현지 시각(stTime). 관리자가 매 스캔 채움
END_VAR
SUPER^.M_Enter(i_stView := i_stView);
_tonRun(IN := FALSE);		// 운전 시간을 처음부터 셈
END_METHOD

METHOD M_Calc : ST_CtrlModeOut
VAR_INPUT
	i_stView	: ST_CtrlModeView;	// 그룹 값(stGroup)·현지 시각(stTime). 관리자가 매 스캔 채움
END_VAR
_tonRun(IN := i_stSet.tDuration > T#0S, PT := i_stSet.tDuration);
M_Calc.bPSetActive	:= TRUE;
M_Calc.fPSet		:= i_stSet.fPSet;
M_Calc.bQSetActive	:= i_stSet.bQSet;
M_Calc.fQSet		:= i_stSet.fQSet;
M_Calc.bExitReq		:= FALSE;
M_Calc.nReason		:= 0;
IF _tonRun.Q THEN
	M_Calc.bExitReq	:= TRUE;
	M_Calc.nReason	:= RSN_TIME_UP;
END_IF
END_METHOD

METHOD M_CheckSet : WSTRING(63)		// 설정 점검: P·Q가 숫자인지 [결함 13 수정 2026-11-04: 추가. 원래 이 FB에는 점검 없음(바탕 FB 빈 문구)]
M_CheckSet := SUPER^.M_CheckSet();
IF M_CheckSet = "" AND NOT (F_RealOk(i_stSet.fPSet) AND F_RealOk(i_stSet.fQSet)) THEN
	M_CheckSet := "정출력: P·Q 값 숫자 아님";
END_IF
END_METHOD

METHOD M_ReasonText : WSTRING(63)
VAR_INPUT
	i_nReason	: UINT;
END_VAR
CASE i_nReason OF
	RSN_NO_UNIT:	M_ReasonText := "정출력: 가용 유닛 없음";
	RSN_TIME_UP:	M_ReasonText := "정출력: 운전 시간 끝";
ELSE
	M_ReasonText := WCONCAT("이유 ", TO_WSTRING(i_nReason));
END_CASE
END_METHOD

END_FUNCTION_BLOCK

// ---- 99_Test/PRG_TestSchedLive.TcPOU
PROGRAM PRG_TestSchedLive		// 스케줄 모드 실제 경로 시험 (시험 모드, MAIN이 부름): 지금 PLC 시각으로 시간표를 넣고 Auto → 배터리 투입 → Run → 스케줄 모드
// bStart := TRUE로 시작. 충전 칸 -200 kW (지금 분 ~ +2분) → 방전 칸 +100 kW (+2 ~ +4분) → 칸 없음 0 kW. 구간마다 5 s 안정 뒤 가상 PCS 실제 출력을 판정
// PCS1(유닛 1, 관리자 g_fbCtrlMode1)로 시험. 접속점은 실측 그대로(ePccShare := Actual)로 둠 (PCS2는 Manual 0)
// 시험 동안만: 방전 허용 시간 끔 (PLC 시계가 UTC), 가상신호로 수전 500 kW (가상 계측기는 부하가 없어 역송 방지에 걸림). 끝나면 설정·모드를 되돌리고 PCS 정지
VAR
	bStart		: BOOL;				// TRUE로 쓰면 시작 (시작하면 FALSE로 돌아감)
	bDone		: BOOL;				// 끝 (bPass로 결과)
	bPass		: BOOL;				// 세 구간 모두 맞음
	nStep		: UINT;
	wsStep		: WSTRING(80);		// 지금 단계
	wsFail		: WSTRING(80);		// 실패 이유
	(* 넣은 시간표 *)
	nSeason		: UINT;				// 0 여름, 1 봄·가을, 2 겨울
	nDow		: UINT;				// 0 = 일요일
	nChgStart	: UINT;				// HHMM, 충전 칸 시작
	nChgEnd		: UINT;				// HHMM, 충전 칸 끝 = 방전 칸 시작
	nDisEnd		: UINT;				// HHMM, 방전 칸 끝
	(* 지금 값 *)
	stNow		: ST_LocalTime;		// PLC 시각 (MAIN.fbClock)
	nActiveMode	: UINT;				// 관리자 켜진 모드 (2 = 스케줄)
	nSlot		: UINT;				// 스케줄 모드가 맞춘 칸
	nSchedState	: UINT;				// 스케줄 모드 상태 (GVL_CM_RSN)
	fSchedP		: REAL;				// 스케줄 모드가 낸 값 (kW, 방전 +)
	fMgrP		: REAL;				// 관리자 지령 (지령원 출력, kW)
	fUnitP		: REAL;				// 가상 PCS 실제 출력 (kW, 방전 +)
	eRun		: E_RunState;		// 가상 PCS 운전 상태
	(* 판정: 구간마다 안정 뒤 값 *)
	fChgP		: REAL;
	fDisP		: REAL;
	fZeroP		: REAL;
	bChgOk		: BOOL;
	bDisOk		: BOOL;
	bZeroOk		: BOOL;
	(* 내부 *)
	nLastStep	: UINT;
	tonStep		: TON;				// 단계 시간 초과
	tonSettle	: TON;				// 구간 진입 뒤 안정
	bBackedUp	: BOOL;
	stSchedBak	: ST_CmScheduleSet;
	stCommonBak	: ST_CmCommonSet;
	stCmBak		: ST_CtrlModeSet;
	stVirtBak	: ST_VirtualSet;
	stMgrOut	: ST_SourceOutput;
	nMin		: UINT;
	k			: UINT;
END_VAR

// 지금 값 (화면용)
stNow		:= MAIN.fbClock.q_stTime;
nActiveMode	:= GVL_SITE.g_fbCtrlMode1.q_nActive;
nSlot		:= GVL_SITE.g_fbCmSchedule1.q_nSlot;
nSchedState	:= GVL_SITE.g_fbCmSchedule1.q_nState;
fSchedP		:= GVL_SITE.g_fbCmSchedule1.q_fOutP;
stMgrOut	:= GVL_SITE.g_fbCtrlMode1.Output;
fMgrP		:= stMgrOut.fPSet;	// [16번 수정 2026-11-09: 관리자가 접속점 그룹 단위 → 접속점 그룹 지령 칸. 원래 stMgrOut.astUnit[1].fPSet (PCS2는 Manual이라 접속점 그룹 지령이 유닛 1로 감)]
fUnitP		:= MAIN.fbSnapshot.q_astUnit[1].stP.fValue;
eRun		:= MAIN.fbSnapshot.q_astUnit[1].eRunState;

tonStep(IN := nStep >= 20 AND nStep < 90, PT := T#200S);

CASE nStep OF
	0:
		IF bStart THEN
			bStart		:= FALSE;
			bDone		:= FALSE;
			bPass		:= FALSE;
			bChgOk		:= FALSE;
			bDisOk		:= FALSE;
			bZeroOk		:= FALSE;
			fChgP		:= 0.0;
			fDisP		:= 0.0;
			fZeroP		:= 0.0;
			wsFail		:= "";
			nStep		:= 10;
		ELSIF NOT bDone THEN
			wsStep := "대기: bStart := TRUE로 시작";
		END_IF

	10:	// 지금 시각으로 시간표 넣기
		wsStep := "시간표 넣는 중";
		IF NOT stNow.bValid OR stNow.nMonth < 1 OR stNow.nMonth > 12 OR stNow.nDay < 1 OR stNow.nDay > 31 OR stNow.nDayOfWeek > 6 THEN
			wsFail	:= "PLC 시각 무효";
			nStep	:= 90;
		ELSE
			nMin := stNow.nHour * 60 + stNow.nMinute;
			IF nMin + 4 >= 1440 THEN
				wsFail	:= "자정 직전이라 시험 안 함 (몇 분 뒤 다시)";
				nStep	:= 90;
			ELSE
				stSchedBak	:= GVL_PERSIST.g_stModuleSet.stCmSchedule1;
				stCommonBak	:= GVL_PERSIST.g_stModuleSet.stCmCommon;
				stVirtBak	:= GVL_TEST.g_astVirtual[1];
				stCmBak		:= GVL_PERSIST.g_stModuleSet.stCtrlMode1;
				GVL_PERSIST.g_stModuleSet.stCtrlMode1.ePccShare := E_PccShare.Actual;
				bBackedUp	:= TRUE;
				nSeason := GVL_PERSIST.g_stModuleSet.stCmCommon.anSeasonOfMonth[stNow.nMonth];
				IF nSeason > 2 THEN
					nSeason := 0;
				END_IF
				nDow		:= stNow.nDayOfWeek;
				nChgStart	:= (nMin / 60) * 100 + nMin MOD 60;
				nChgEnd		:= ((nMin + 2) / 60) * 100 + (nMin + 2) MOD 60;
				nDisEnd		:= ((nMin + 4) / 60) * 100 + (nMin + 4) MOD 60;
				FOR k := 1 TO GVL_PARAM.SCHED_SLOT_COUNT DO
					GVL_PERSIST.g_stModuleSet.stCmSchedule1.astSlot[nSeason, nDow, k].nStart	:= 0;
					GVL_PERSIST.g_stModuleSet.stCmSchedule1.astSlot[nSeason, nDow, k].nEnd	:= 0;
					GVL_PERSIST.g_stModuleSet.stCmSchedule1.astSlot[nSeason, nDow, k].fP		:= 0.0;
				END_FOR
				GVL_PERSIST.g_stModuleSet.stCmSchedule1.astSlot[nSeason, nDow, 1].nStart	:= nChgStart;
				GVL_PERSIST.g_stModuleSet.stCmSchedule1.astSlot[nSeason, nDow, 1].nEnd	:= nChgEnd;
				GVL_PERSIST.g_stModuleSet.stCmSchedule1.astSlot[nSeason, nDow, 1].fP		:= -200.0;
				GVL_PERSIST.g_stModuleSet.stCmSchedule1.astSlot[nSeason, nDow, 2].nStart	:= nChgEnd;
				GVL_PERSIST.g_stModuleSet.stCmSchedule1.astSlot[nSeason, nDow, 2].nEnd	:= nDisEnd;
				GVL_PERSIST.g_stModuleSet.stCmSchedule1.astSlot[nSeason, nDow, 2].fP		:= 100.0;
				GVL_PERSIST.g_stModuleSet.stCmCommon.abHoliday[stNow.nMonth, stNow.nDay]	:= FALSE;
				GVL_PERSIST.g_stModuleSet.stCmCommon.stDis.bUse	:= FALSE;
				GVL_TEST.g_astVirtual[1].bPEna	:= TRUE;
				GVL_TEST.g_astVirtual[1].fP		:= -500.0;		// 수전 500 kW
				GVL_PERSIST.g_aeOpMode[1]		:= E_OpMode.Auto;
				nStep := 20;
			END_IF
		END_IF

	20:	// Auto 전환 → 배터리 투입 요청
		wsStep := "Auto 전환 대기";
		IF MAIN.fbModeSwitch.q_aeOpMode[1] = E_OpMode.Auto THEN
			GVL_SITE.g_fbSrcTest.i_nBatGroup	:= 0;
			GVL_SITE.g_fbSrcTest.i_eBatReq		:= E_BatCmd.Close;
			nStep := 30;
		END_IF

	30:	// 배터리 투입 → Run 요청
		wsStep := "배터리 투입 대기";
		IF MAIN.fbBatGroup.q_astBatGroup[1].bReady THEN
			GVL_SITE.g_fbSrcTest.i_nPcsUnit	:= 0;
			GVL_SITE.g_fbSrcTest.i_ePcsReq	:= E_PcsCmd.Run;
			nStep := 40;
		END_IF

	40:	// Run → 스케줄 모드(2) 요청
		wsStep := "PCS Run 대기";
		IF eRun = E_RunState.Run THEN
			GVL_SITE.g_fbCtrlMode1.i_nModeReq := 2;
			nStep := 50;
		END_IF

	50:
		wsStep := "스케줄 모드 켜는 중";
		IF nActiveMode = 2 THEN
			nStep := 60;
		END_IF

	60:	// 충전 칸
		wsStep := "충전 칸: -200 kW";
		tonSettle(IN := nSlot = 1, PT := T#5S);
		IF tonSettle.Q THEN
			fChgP	:= fUnitP;
			bChgOk	:= ABS(fUnitP + 200.0) < 5.0 AND ABS(fSchedP + 200.0) < 0.1 AND ABS(fMgrP + 200.0) < 0.1;
		END_IF
		IF nSlot = 2 THEN
			tonSettle(IN := FALSE);
			nStep := 70;
		END_IF

	70:	// 방전 칸
		wsStep := "방전 칸: +100 kW";
		tonSettle(IN := nSlot = 2, PT := T#5S);
		IF tonSettle.Q THEN
			fDisP	:= fUnitP;
			bDisOk	:= ABS(fUnitP - 100.0) < 5.0 AND ABS(fSchedP - 100.0) < 0.1 AND ABS(fMgrP - 100.0) < 0.1;
		END_IF
		IF nSlot = 0 THEN
			tonSettle(IN := FALSE);
			nStep := 80;
		END_IF

	80:	// 칸 없음 → 0
		wsStep := "칸 없음: 0 kW";
		tonSettle(IN := nSlot = 0, PT := T#5S);
		IF tonSettle.Q THEN
			fZeroP	:= fUnitP;
			bZeroOk	:= ABS(fUnitP) < 5.0 AND nSchedState = GVL_CM_RSN.NO_SLOT AND stMgrOut.bPSetActive;	// [16번 수정 2026-11-09: 원래 stMgrOut.astUnit[1].bPSetActive]
			tonSettle(IN := FALSE);
			nStep := 90;
		END_IF

	90:	// 정리: 모드 끔, PCS 정지, 설정·가상신호·운전 모드 되돌림
		GVL_SITE.g_fbCtrlMode1.i_nModeReq	:= 0;
		GVL_SITE.g_fbSrcTest.i_nPcsUnit		:= 0;
		GVL_SITE.g_fbSrcTest.i_ePcsReq		:= E_PcsCmd.Stop;
		IF bBackedUp THEN
			GVL_PERSIST.g_stModuleSet.stCmSchedule1	:= stSchedBak;
			GVL_PERSIST.g_stModuleSet.stCmCommon	:= stCommonBak;
			GVL_TEST.g_astVirtual[1]				:= stVirtBak;
			GVL_PERSIST.g_stModuleSet.stCtrlMode1	:= stCmBak;
			bBackedUp := FALSE;
		END_IF
		GVL_PERSIST.g_aeOpMode[1] := E_OpMode.Manual;
		bPass	:= bChgOk AND bDisOk AND bZeroOk AND wsFail = "";
		bDone	:= TRUE;
		IF bPass THEN
			wsStep := "끝: 통과";
		ELSE
			wsStep := "끝: 실패 (wsFail·구간 값 확인)";
		END_IF
		nStep := 0;
END_CASE

// 단계 시간 초과
IF tonStep.Q AND nStep >= 20 AND nStep < 90 THEN
	wsFail	:= WCONCAT("시간 초과: ", wsStep);
	nStep	:= 90;
END_IF
IF nStep <> nLastStep THEN
	tonStep(IN := FALSE);
	nLastStep := nStep;
END_IF

END_PROGRAM

// ---- 99_Test/PRG_TestPeakLive.TcPOU
PROGRAM PRG_TestPeakLive		// 피크컷(3)·통합(4) 모드 실제 경로 시험 (시험 모드, MAIN이 부름). bStart := TRUE로 시작, 약 10~15분
// 부하 모델: 가상 접속점 P = ESS 출력 − 부하 (수전 = 부하 − ESS 방전). 목표 피크 300 kW, 방전 허용 시간 끔 (PLC 시계 UTC)
// 피크컷: P1 부하 500 → 피크 방전, P2 부하 200 → 0, P3 자동 충전 시간 → 충전, P4 잔량 방전 시간 → 방전 (역송 방지 상한)
// 통합:   I1 부하 200·시간표 +100 → 100, I2 부하 600 → 피크·시간표 중 큰 값, I3 부하 200·시간표 −200 → 충전, I4 잔량 방전
// 구간마다 조건이 5 s 이어지면 통과·기록. 끝나면 설정·가상신호·운전 모드 되돌리고 PCS 정지
VAR
	bStart		: BOOL;				// TRUE로 쓰면 시작
	bDone		: BOOL;
	bPass		: BOOL;				// 8구간 모두 통과
	nStep		: UINT;
	wsStep		: WSTRING(80);		// 지금 단계
	wsFail		: WSTRING(80);
	(* 지금 값 *)
	fLoadSim	: REAL;				// kW, 모의 부하
	fImport		: REAL;				// kW, 수전 (= 부하 − ESS 출력)
	nActiveMode	: UINT;				// 3 = 피크컷, 4 = 통합
	nState		: UINT;				// 켜진 모드 상태 (GVL_CM_RSN: 0 정상, 11 피크, 12 피크 필요 없음, 13 자동 충전, 14 잔량 방전, 15 스케줄·피크, 6 역송 방지)
	fModeP		: REAL;				// 모드가 낸 값 (kW, 방전 +)
	fMgrP		: REAL;				// 관리자 지령
	fUnitP		: REAL;				// 가상 PCS 실제 출력
	fPeakCtrl	: REAL;				// 피크 제어량
	nRemainMin	: UINT;				// 15분 구간 남은 분
	fSoc		: REAL;				// %
	eRun		: E_RunState;
	stNow		: ST_LocalTime;
	(* 구간 결과 (통과 때 실제 출력 kW) *)
	bP1Peak		: BOOL;		fP1		: REAL;		// 피크컷: 부하 500 → 피크 방전
	bP2Below	: BOOL;		fP2		: REAL;		// 피크컷: 부하 200 → 0
	bP3AutoChg	: BOOL;		fP3		: REAL;		// 피크컷: 자동 충전
	bP4Remain	: BOOL;		fP4		: REAL;		// 피크컷: 잔량 방전
	bI1Sched	: BOOL;		fI1		: REAL;		// 통합: 시간표 +100
	bI2Peak		: BOOL;		fI2		: REAL;		// 통합: 피크·시간표 중 큰 값
	bI3Chg		: BOOL;		fI3		: REAL;		// 통합: 시간표 충전 −200
	bI4Remain	: BOOL;		fI4		: REAL;		// 통합: 잔량 방전
	(* 내부 *)
	bLoadSim	: BOOL;
	nLastStep	: UINT;
	tonStep		: TON;
	tonOk		: TON;
	bCond		: BOOL;
	bBackedUp	: BOOL;
	stCommonBak	: ST_CmCommonSet;
	stSchedBak	: ST_CmScheduleSet;
	stPeakBak	: ST_CmPeakCutSet;
	stSPBak		: ST_CmSchedPeakSet;
	stVirtBak	: ST_VirtualSet;
	stCmBak		: ST_CtrlModeSet;
	stMgrOut	: ST_SourceOutput;
	nMin		: UINT;
	nSeason		: UINT;
	k			: UINT;
	nWinStart	: UINT;		// HHMM
	nWinEnd		: UINT;		// HHMM (지금 + 3분)
	nSlotEnd	: UINT;		// HHMM (지금 + 30분)
END_VAR

// 지금 값
stNow		:= MAIN.fbClock.q_stTime;
nActiveMode	:= GVL_SITE.g_fbCtrlMode1.q_nActive;
stMgrOut	:= GVL_SITE.g_fbCtrlMode1.Output;
fMgrP		:= stMgrOut.fPSet;	// [16번 수정 2026-11-09: 관리자가 접속점 그룹 단위 → 접속점 그룹 지령 칸. 원래 stMgrOut.astUnit[1].fPSet (PCS2는 Manual이라 접속점 그룹 지령이 유닛 1로 감)]
fUnitP		:= MAIN.fbSnapshot.q_astUnit[1].stP.fValue;
eRun		:= MAIN.fbSnapshot.q_astUnit[1].eRunState;
fSoc		:= MAIN.fbGroupView.q_astView[1].stSocAvg.fValue;
IF nActiveMode = 4 THEN
	nState		:= GVL_SITE.g_fbCmSchedPeak1.q_nState;
	fModeP		:= GVL_SITE.g_fbCmSchedPeak1.q_fOutP;
	fPeakCtrl	:= GVL_SITE.g_fbCmSchedPeak1.q_fPeakCtrl;
	nRemainMin	:= GVL_SITE.g_fbCmSchedPeak1.q_nRemainMin;
ELSE
	nState		:= GVL_SITE.g_fbCmPeakCut1.q_nState;
	fModeP		:= GVL_SITE.g_fbCmPeakCut1.q_fOutP;
	fPeakCtrl	:= GVL_SITE.g_fbCmPeakCut1.q_fPeakCtrl;
	nRemainMin	:= GVL_SITE.g_fbCmPeakCut1.q_nRemainMin;
END_IF
// 부하 모델: 접속점 P (공급 +) = ESS 출력 − 부하
IF bLoadSim THEN
	GVL_TEST.g_astVirtual[1].bPEna	:= TRUE;
	GVL_TEST.g_astVirtual[1].fP		:= MAIN.fbGroupView.q_astView[1].fPOut - fLoadSim;	// 그룹 출력 (PCS2는 Manual 0)
END_IF
fImport := fLoadSim - fUnitP;
// 시간 구간 (지금 분 ~ +3분, 시간표 칸은 +30분)
nMin		:= stNow.nHour * 60 + stNow.nMinute;
nWinStart	:= (nMin / 60) * 100 + nMin MOD 60;
nWinEnd		:= (((nMin + 3) MOD 1440) / 60) * 100 + ((nMin + 3) MOD 1440) MOD 60;
nSlotEnd	:= (((nMin + 30) MOD 1440) / 60) * 100 + ((nMin + 30) MOD 1440) MOD 60;

tonStep(IN := nStep >= 20 AND nStep < 900, PT := T#240S);
bCond := FALSE;

CASE nStep OF
	0:
		IF bStart THEN
			bStart := FALSE;	bDone := FALSE;	bPass := FALSE;	wsFail := "";
			bP1Peak := FALSE;	bP2Below := FALSE;	bP3AutoChg := FALSE;	bP4Remain := FALSE;
			bI1Sched := FALSE;	bI2Peak := FALSE;	bI3Chg := FALSE;	bI4Remain := FALSE;
			nStep := 10;
		ELSIF NOT bDone THEN
			wsStep := "대기: bStart := TRUE로 시작";
		END_IF

	10:	// 준비
		wsStep := "설정 준비";
		IF NOT stNow.bValid OR stNow.nMonth < 1 OR stNow.nMonth > 12 OR stNow.nDay < 1 OR stNow.nDay > 31 OR stNow.nDayOfWeek > 6 THEN
			wsFail := "PLC 시각 무효";
			nStep := 900;
		ELSIF nMin + 40 >= 1440 THEN
			wsFail := "자정 가까움: 40분 뒤 다시";
			nStep := 900;
		ELSE
			stCommonBak	:= GVL_PERSIST.g_stModuleSet.stCmCommon;
			stSchedBak	:= GVL_PERSIST.g_stModuleSet.stCmSchedule1;
			stPeakBak	:= GVL_PERSIST.g_stModuleSet.stCmPeakCut1;
			stSPBak		:= GVL_PERSIST.g_stModuleSet.stCmSchedPeak1;
			stVirtBak	:= GVL_TEST.g_astVirtual[1];
			stCmBak		:= GVL_PERSIST.g_stModuleSet.stCtrlMode1;
			GVL_PERSIST.g_stModuleSet.stCtrlMode1.ePccShare := E_PccShare.Actual;	// PCS1이 접속점 실측 그대로 (PCS2는 Manual 0)
			bBackedUp	:= TRUE;
			GVL_PERSIST.g_stModuleSet.stCmCommon.stDis.bUse := FALSE;
			GVL_PERSIST.g_stModuleSet.stCmCommon.abHoliday[stNow.nMonth, stNow.nDay] := FALSE;
			GVL_PERSIST.g_stModuleSet.stCmPeakCut1.stPeak.fTarget	:= 300.0;
			GVL_PERSIST.g_stModuleSet.stCmPeakCut1.stAutoChg.bUse	:= FALSE;
			GVL_PERSIST.g_stModuleSet.stCmPeakCut1.stRemain.bUse		:= FALSE;
			GVL_PERSIST.g_stModuleSet.stCmSchedPeak1.stPeak.fTarget	:= 300.0;
			GVL_PERSIST.g_stModuleSet.stCmSchedPeak1.stRemain.bUse	:= FALSE;
			nSeason := GVL_PERSIST.g_stModuleSet.stCmCommon.anSeasonOfMonth[stNow.nMonth];
			IF nSeason > 2 THEN
				nSeason := 0;
			END_IF
			FOR k := 1 TO GVL_PARAM.SCHED_SLOT_COUNT DO
				GVL_PERSIST.g_stModuleSet.stCmSchedule1.astSlot[nSeason, stNow.nDayOfWeek, k].nStart	:= 0;
				GVL_PERSIST.g_stModuleSet.stCmSchedule1.astSlot[nSeason, stNow.nDayOfWeek, k].nEnd	:= 0;
				GVL_PERSIST.g_stModuleSet.stCmSchedule1.astSlot[nSeason, stNow.nDayOfWeek, k].fP		:= 0.0;
			END_FOR
			fLoadSim	:= 500.0;
			bLoadSim	:= TRUE;
			GVL_PERSIST.g_aeOpMode[1] := E_OpMode.Auto;
			nStep := 20;
		END_IF

	20:
		wsStep := "Auto 전환 대기";
		IF MAIN.fbModeSwitch.q_aeOpMode[1] = E_OpMode.Auto THEN
			GVL_SITE.g_fbSrcTest.i_nBatGroup	:= 0;
			GVL_SITE.g_fbSrcTest.i_eBatReq		:= E_BatCmd.Close;
			nStep := 30;
		END_IF
	30:
		wsStep := "배터리 투입 대기";
		IF MAIN.fbBatGroup.q_astBatGroup[1].bReady THEN
			GVL_SITE.g_fbSrcTest.i_nPcsUnit	:= 0;
			GVL_SITE.g_fbSrcTest.i_ePcsReq	:= E_PcsCmd.Run;
			nStep := 40;
		END_IF
	40:
		wsStep := "PCS Run 대기";
		IF eRun = E_RunState.Run THEN
			GVL_SITE.g_fbCtrlMode1.i_nModeReq := 3;
			nStep := 50;
		END_IF
	50:
		wsStep := "피크컷 모드 켜는 중";
		IF nActiveMode = 3 THEN
			nStep := 100;
		END_IF

	100: // P1 부하 500 > 목표 300 → 피크 방전
		wsStep := "P1 피크컷: 부하 500 > 목표 300";
		bCond := nActiveMode = 3 AND nState = GVL_CM_RSN.PEAK AND fPeakCtrl > 0.0 AND fModeP > 0.0 AND ABS(fUnitP - fModeP) < 5.0;
		IF tonOk.Q THEN
			bP1Peak := TRUE;	fP1 := fUnitP;
			fLoadSim := 200.0;
			nStep := 110;
		END_IF
	110: // P2 부하 200 < 목표 → 0
		wsStep := "P2 피크컷: 부하 200 < 목표 300";
		bCond := nState = GVL_CM_RSN.BELOW_PEAK AND ABS(fUnitP) < 5.0;
		IF tonOk.Q THEN
			bP2Below := TRUE;	fP2 := fUnitP;
			GVL_PERSIST.g_stModuleSet.stCmPeakCut1.stAutoChg.nStart	:= nWinStart;
			GVL_PERSIST.g_stModuleSet.stCmPeakCut1.stAutoChg.nEnd	:= nWinEnd;
			GVL_PERSIST.g_stModuleSet.stCmPeakCut1.stAutoChg.fSoc	:= 100.0;
			GVL_PERSIST.g_stModuleSet.stCmPeakCut1.stAutoChg.bUse	:= TRUE;
			nStep := 120;
		END_IF
	120: // P3 자동 충전 시간
		wsStep := "P3 피크컷: 자동 충전 시간";
		bCond := nState = GVL_CM_RSN.AUTO_CHG AND fModeP < -5.0 AND fUnitP < -5.0;
		IF tonOk.Q THEN
			bP3AutoChg := TRUE;	fP3 := fUnitP;
			GVL_PERSIST.g_stModuleSet.stCmPeakCut1.stAutoChg.bUse	:= FALSE;
			GVL_PERSIST.g_stModuleSet.stCmPeakCut1.stRemain.nStart	:= nWinStart;
			GVL_PERSIST.g_stModuleSet.stCmPeakCut1.stRemain.nEnd		:= nWinEnd;
			GVL_PERSIST.g_stModuleSet.stCmPeakCut1.stRemain.fSoc		:= 10.0;
			GVL_PERSIST.g_stModuleSet.stCmPeakCut1.stRemain.bUse		:= TRUE;
			fLoadSim := 500.0;
			nStep := 130;
		END_IF
	130: // P4 잔량 방전 시간 (역송 방지 상한)
		wsStep := "P4 피크컷: 잔량 방전 시간";
		bCond := (nState = GVL_CM_RSN.REMAIN_DIS OR nState = GVL_CM_RSN.REV_LIMIT) AND fModeP > 5.0 AND ABS(fUnitP - fModeP) < 5.0 AND fUnitP < fLoadSim;
		IF tonOk.Q THEN
			bP4Remain := TRUE;	fP4 := fUnitP;
			GVL_PERSIST.g_stModuleSet.stCmPeakCut1.stRemain.bUse := FALSE;
			// 통합 준비: 시간표 +100 (지금 ~ +30분), 부하 200
			GVL_PERSIST.g_stModuleSet.stCmSchedule1.astSlot[nSeason, stNow.nDayOfWeek, 1].nStart	:= nWinStart;
			GVL_PERSIST.g_stModuleSet.stCmSchedule1.astSlot[nSeason, stNow.nDayOfWeek, 1].nEnd	:= nSlotEnd;
			GVL_PERSIST.g_stModuleSet.stCmSchedule1.astSlot[nSeason, stNow.nDayOfWeek, 1].fP		:= 100.0;
			fLoadSim := 200.0;
			GVL_SITE.g_fbCtrlMode1.i_nModeReq := 4;
			nStep := 200;
		END_IF

	200:
		wsStep := "통합 모드 켜는 중";
		IF nActiveMode = 4 THEN
			nStep := 210;
		END_IF
	210: // I1 부하 200 (피크 아님) → 시간표 +100
		wsStep := "I1 통합: 부하 200, 시간표 +100";
		bCond := nState = 0 AND ABS(fModeP - 100.0) < 0.5 AND ABS(fUnitP - 100.0) < 5.0;
		IF tonOk.Q THEN
			bI1Sched := TRUE;	fI1 := fUnitP;
			fLoadSim := 600.0;
			nStep := 220;
		END_IF
	220: // I2 부하 600 > 목표 → 피크 제어량과 시간표 중 큰 값
		wsStep := "I2 통합: 부하 600 > 목표 300";
		bCond := nState = GVL_CM_RSN.SCHED_PEAK AND fPeakCtrl > 0.0 AND fModeP >= 99.9 AND ABS(fModeP - MAX(fPeakCtrl, 100.0)) < 0.5 AND ABS(fUnitP - fModeP) < 5.0;
		IF tonOk.Q THEN
			bI2Peak := TRUE;	fI2 := fUnitP;
			GVL_PERSIST.g_stModuleSet.stCmSchedule1.astSlot[nSeason, stNow.nDayOfWeek, 1].fP := -200.0;
			fLoadSim := 200.0;
			nStep := 230;
		END_IF
	230: // I3 부하 200, 시간표 충전 −200
		wsStep := "I3 통합: 부하 200, 시간표 -200";
		bCond := nState = 0 AND ABS(fModeP + 200.0) < 0.5 AND ABS(fUnitP + 200.0) < 5.0;
		IF tonOk.Q THEN
			bI3Chg := TRUE;	fI3 := fUnitP;
			GVL_PERSIST.g_stModuleSet.stCmSchedPeak1.stRemain.nStart	:= nWinStart;
			GVL_PERSIST.g_stModuleSet.stCmSchedPeak1.stRemain.nEnd	:= nWinEnd;
			GVL_PERSIST.g_stModuleSet.stCmSchedPeak1.stRemain.fSoc	:= 10.0;
			GVL_PERSIST.g_stModuleSet.stCmSchedPeak1.stRemain.bUse	:= TRUE;
			fLoadSim := 500.0;
			nStep := 240;
		END_IF
	240: // I4 잔량 방전
		wsStep := "I4 통합: 잔량 방전 시간";
		bCond := (nState = GVL_CM_RSN.REMAIN_DIS OR nState = GVL_CM_RSN.REV_LIMIT) AND fModeP > 5.0 AND ABS(fUnitP - fModeP) < 5.0 AND fUnitP < fLoadSim;
		IF tonOk.Q THEN
			bI4Remain := TRUE;	fI4 := fUnitP;
			nStep := 900;
		END_IF

	900: // 정리
		GVL_SITE.g_fbCtrlMode1.i_nModeReq	:= 0;
		GVL_SITE.g_fbSrcTest.i_nPcsUnit		:= 0;
		GVL_SITE.g_fbSrcTest.i_ePcsReq		:= E_PcsCmd.Stop;
		bLoadSim := FALSE;
		IF bBackedUp THEN
			GVL_PERSIST.g_stModuleSet.stCmCommon	:= stCommonBak;
			GVL_PERSIST.g_stModuleSet.stCmSchedule1	:= stSchedBak;
			GVL_PERSIST.g_stModuleSet.stCmPeakCut1	:= stPeakBak;
			GVL_PERSIST.g_stModuleSet.stCmSchedPeak1	:= stSPBak;
			GVL_TEST.g_astVirtual[1]				:= stVirtBak;
			GVL_PERSIST.g_stModuleSet.stCtrlMode1	:= stCmBak;
			bBackedUp := FALSE;
		END_IF
		GVL_PERSIST.g_aeOpMode[1] := E_OpMode.Manual;
		bPass := bP1Peak AND bP2Below AND bP3AutoChg AND bP4Remain AND bI1Sched AND bI2Peak AND bI3Chg AND bI4Remain AND wsFail = "";
		bDone := TRUE;
		IF bPass THEN
			wsStep := "끝: 통과";
		ELSE
			wsStep := "끝: 실패 (wsFail·구간 결과 확인)";
		END_IF
		nStep := 0;
END_CASE

// 조건이 5 s 이어지면 통과 (단계가 바뀌면 다시 셈)
tonOk(IN := bCond AND nStep = nLastStep, PT := T#5S);
IF tonStep.Q AND nStep >= 20 AND nStep < 900 THEN
	wsFail	:= WCONCAT("시간 초과: ", wsStep);
	nStep	:= 900;
END_IF
IF nStep <> nLastStep THEN
	tonStep(IN := FALSE);
	tonOk(IN := FALSE);
	nLastStep := nStep;
END_IF

END_PROGRAM

// ---- 99_Test/PRG_TestUnitMode.TcPOU
PROGRAM PRG_TestUnitMode		// PCS별(유닛 단위) 제어 모드 자동 시험 (GVL_SITE.TEST_MODE일 때 MAIN이 부름). 따로 둔 인스턴스만 씀 (장비 지령에 영향 없음)
// 온라인에서 bDone = TRUE가 되면 fbTally.q_nPass·q_nFail, 실패하면 fbTally.q_anFail. bRestart := TRUE로 다시 돌림
// 40~41: 유닛 단위 출력 칸, 42~44: 접속점 몫 (ByRating·Actual·Fixed), 45~47: 설정 점검, 48~50: FB_UnitView 버스 몫, 51~57: 스탠다드 스케줄 모드, 58~63: NaN·무한대 거르기 (PLC가 멈추지 않아야 함)
VAR
	bRestart	: BOOL;
	bDone		: BOOL;
	nStep		: UINT;
	fbTally		: FB_TestTally;
	fbConstU	: FB_CmConstPower	:= (i_nModuleId := 9012, i_sName := 'TestConstU');
	fbMgrU		: FB_CtrlModeMgr	:= (i_nModuleId := 9010, i_sName := 'TestMgrU', i_nUnit := 1);
	aipMode		: ARRAY[1..GVL_PARAM.CTRL_MODE_COUNT] OF I_ControlMode;
	astUv		: ARRAY[1..GVL_PARAM.UNIT_COUNT] OF ST_UnitView;	// 관리자에 주소로 넘기는 유닛 값 (시험이 채움)
	stGrpView	: ST_GroupView;			// 지령원 공통 입력 (유닛 단위에서는 안 봄)
	stReg		: ST_SourceReg := (bEnable := TRUE, nGrade := 1, ePowerMode := E_SourceMode.Auto, nGroup := 0, tExpire := T#10S);
	stMgrOut	: ST_SourceOutput;
	wsTmp		: WSTRING(63);
	(* FB_UnitView 시험 (유닛 1 기준, 유닛이 2개 이상이면 유닛 2도) *)
	fbUv		: FB_UnitView;
	astView		: ARRAY[1..GVL_PARAM.GROUP_COUNT] OF ST_GroupView;
	astUnit		: ARRAY[1..GVL_PARAM.UNIT_COUNT] OF ST_UnitState;
	astAvail	: ARRAY[1..GVL_PARAM.UNIT_COUNT] OF ST_UnitAvail;
	astCfg		: ARRAY[1..GVL_PARAM.UNIT_COUNT] OF ST_UnitCfg;
	astEnv		: ARRAY[1..GVL_PARAM.UNIT_COUNT] OF ST_UnitEnvelope;
	astBat		: ARRAY[1..GVL_PARAM.BAT_COUNT] OF ST_BatGroupState;
	astBatEnv	: ARRAY[1..GVL_PARAM.BAT_COUNT] OF ST_BatEnvelope;
	fShareExp	: REAL;
	(* 스탠다드 스케줄 모드 시험 *)
	fbStd		: FB_CmStdSchedule	:= (i_nModuleId := 9013, i_sName := 'TestStdSched');
	stStdView	: ST_CtrlModeView;
	stStdOut	: ST_CtrlModeOut;
	nInfBits	: DWORD := 16#7F800000;	// +무한대 비트 (NaN은 크기 비교에서 부동소수점 예외로 PLC가 멈추므로 시험에 쓰지 않음)
	fInf		: REAL;
	nBad0		: UDINT;
	nNanBits	: DWORD := 16#7FC00000;	// NaN 비트 (거르기 시험: 비교하기 전에 걸러져야 PLC가 멈추지 않음)
	fNan		: REAL;
	fbEmsCmd	: FB_EmsCommand;		// EMS 명령 핸들러 시험 인스턴스
	astPcsRx	: ARRAY[0..GVL_PARAM.PCS_COUNT - 1] OF ST_MqttCommand_Rx;
	astBatRx	: ARRAY[0..GVL_PARAM.BMS_COUNT - 1] OF ST_MqttCommand_Rx;
	nPSeq0		: UDINT;
	nRunSeq0	: UDINT;		// 시험 전 이상값 버린 수 (누계라 다시 돌려도 맞게)
	u			: UINT;
END_VAR

IF bRestart THEN
	bRestart	:= FALSE;
	bDone		:= FALSE;
	nStep		:= 0;
END_IF

CASE nStep OF
	0:	// 준비: 정출력 80 kW 하나, 유닛 1 값 (출력 100, 그룹 출력 300, 접속점 -200 = 수전 200 → 그룹 부하 500, 몫 0.5)
		fbTally.M_Reset();
		aipMode[1]					:= fbConstU;
		fbConstU.i_stSet.fPSet		:= 80.0;
		fbConstU.i_stSet.bQSet		:= FALSE;
		fbConstU.i_stSet.tDuration	:= T#0S;
		astUv[1].nUnit				:= 1;
		astUv[1].bAvail				:= TRUE;
		astUv[1].stView.nUnitAvail	:= 1;
		astUv[1].stView.fPRatedAvail	:= 1000.0;
		astUv[1].stView.fPOut		:= 100.0;
		astUv[1].stView.stPcc.stMeas.stP.bValid	:= TRUE;
		astUv[1].stView.stPcc.stMeas.stP.fValue	:= -200.0;
		astUv[1].fGroupPOut			:= 300.0;
		astUv[1].fRatingShare		:= 0.5;
		fbMgrU.i_aipMode			:= aipMode;
		fbMgrU.i_stSet.bZeroOnSwitch	:= TRUE;
		fbMgrU.i_stSet.tZeroDelay	:= T#1S;
		fbMgrU.i_stSet.nFallback	:= 0;
		fbMgrU.i_stSet.ePccShare	:= E_PccShare.ByRating;
		fbMgrU.i_stSet.fPccRatio	:= 1.0;
		fbMgrU.i_pUnitView			:= ADR(astUv);
		wsTmp := fbMgrU.M_CheckSet();
		fbTally.M_Check(i_nId := 40, i_bOk := wsTmp = "");
		fbMgrU.i_nModeReq := 1;
		nStep := 10;

	10:	// 정출력 진입: 유닛 1 칸에만 80, 그룹 지령은 없음. 몫 0.5 → 모드가 본 접속점 = 100 - 0.5 × 500 = -150
		A_Cycle();
		fbTally.M_Check(i_nId := 41, i_bOk := fbMgrU.q_nActive = 1 AND stMgrOut.astUnit[1].bPSetActive AND ABS(stMgrOut.astUnit[1].fPSet - 80.0) < 0.01 AND NOT stMgrOut.bPSetActive);
		fbTally.M_Check(i_nId := 42, i_bOk := ABS(fbMgrU.q_fPccP + 150.0) < 0.01);
		fbMgrU.i_stSet.ePccShare := E_PccShare.Actual;
		nStep := 11;

	11:	// Actual: 실측 그대로 -200
		A_Cycle();
		fbTally.M_Check(i_nId := 43, i_bOk := ABS(fbMgrU.q_fPccP + 200.0) < 0.01);
		fbMgrU.i_stSet.ePccShare := E_PccShare.Fixed;
		fbMgrU.i_stSet.fPccRatio := 0.2;
		nStep := 12;

	12:	// Fixed 0.2: 100 - 0.2 × 500 = 0
		A_Cycle();
		fbTally.M_Check(i_nId := 44, i_bOk := ABS(fbMgrU.q_fPccP) < 0.01);
		// 설정 점검: 몫 범위 밖, 유닛 값 연결 안 됨, 유닛 번호 범위 밖
		fbMgrU.i_stSet.fPccRatio := 1.5;
		wsTmp := fbMgrU.M_CheckSet();
		fbTally.M_Check(i_nId := 45, i_bOk := wsTmp <> "");
		fbMgrU.i_stSet.fPccRatio := 0.2;
		fbMgrU.i_pUnitView := 0;
		wsTmp := fbMgrU.M_CheckSet();
		fbTally.M_Check(i_nId := 46, i_bOk := wsTmp <> "");
		fbMgrU.i_pUnitView := ADR(astUv);
		fbMgrU.i_nUnit := GVL_PARAM.UNIT_COUNT + 1;
		wsTmp := fbMgrU.M_CheckSet();
		fbTally.M_Check(i_nId := 47, i_bOk := wsTmp <> "");
		fbMgrU.i_nUnit := 1;
		A_UnitViewTest();
		A_StdScheduleTest();
		A_NanTest();
		nStep := 99;

	99:
		bDone := TRUE;
END_CASE

ACTION A_Cycle:
fbMgrU.i_pUnitView := ADR(astUv);	// 온라인 변경 뒤에도 맞게 매번
fbMgrU.M_Cycle(i_stReg := stReg, i_stView := stGrpView);
stMgrOut := fbMgrU.Output;
END_ACTION

ACTION A_UnitViewTest:
// FB_UnitView: 그룹 1 (접속점 -200, 그룹 출력 300, 가용 한도 합 2000), 버스 1 (방전 한도 1200, 충전 한도 800, 용량 4000, SOC 60)
// 유닛 1 정격 1000 (한도 1000, 출력 100). 유닛이 2개 이상이면 유닛 2도 같은 버스·정격 1000 → 버스 몫 0.5, 아니면 1
astView[1].stPcc.stMeas.stP.bValid	:= TRUE;
astView[1].stPcc.stMeas.stP.fValue	:= -200.0;
astView[1].fPOut			:= 300.0;
astView[1].fPRatedAvail		:= 2000.0;
astBat[1].bUsable			:= TRUE;
astBat[1].fCapacity			:= 4000.0;
astBat[1].stSoc.bValid		:= TRUE;
astBat[1].stSoc.fValue		:= 60.0;
astBatEnv[1].stP.fMax		:= 1200.0;
astBatEnv[1].stP.fMin		:= -800.0;
FOR u := 1 TO GVL_PARAM.UNIT_COUNT DO
	astCfg[u].nGroup		:= 1;
	astCfg[u].nBatGroup		:= 1;
	astCfg[u].fPRated		:= 1000.0;
	astCfg[u].fQRated		:= 500.0;
	astAvail[u].bAvail		:= TRUE;
	astEnv[u].stP.fMax		:= 1000.0;
	astEnv[u].stQ.fMax		:= 500.0;
	astUnit[u].stP.bValid	:= TRUE;
	astUnit[u].stP.fValue	:= 100.0;
END_FOR
fShareExp := 1.0 / UINT_TO_REAL(GVL_PARAM.UNIT_COUNT);
fbUv(iq_astView := astView, iq_astUnit := astUnit, iq_astAvail := astAvail, iq_astUnitCfg := astCfg,
	iq_astUnitEnv := astEnv, iq_astBatGroup := astBat, iq_astBatEnv := astBatEnv);
// 48) 유닛 1: 출력·한도·접속점·그룹 출력·정격 몫 (1000 / 2000)
fbTally.M_Check(i_nId := 48, i_bOk := fbUv.q_astView[1].stView.nUnitAvail = 1 AND ABS(fbUv.q_astView[1].stView.fPOut - 100.0) < 0.01
	AND ABS(fbUv.q_astView[1].stView.fPRatedAvail - 1000.0) < 0.01 AND ABS(fbUv.q_astView[1].stView.stPcc.stMeas.stP.fValue + 200.0) < 0.01
	AND ABS(fbUv.q_astView[1].fGroupPOut - 300.0) < 0.01 AND ABS(fbUv.q_astView[1].fRatingShare - 0.5) < 0.001);
// 49) 버스 몫: 용량·방전·충전 한도 × 몫, SOC 그대로
fbTally.M_Check(i_nId := 49, i_bOk := ABS(fbUv.q_astView[1].stView.fCapacity - 4000.0 * fShareExp) < 0.1
	AND ABS(fbUv.q_astView[1].stView.fPDisMax - MIN(1200.0 * fShareExp, 1000.0)) < 0.1 AND ABS(fbUv.q_astView[1].stView.fPChgMax - MIN(800.0 * fShareExp, 1000.0)) < 0.1
	AND fbUv.q_astView[1].stView.stSocAvg.bValid AND ABS(fbUv.q_astView[1].stView.stSocAvg.fValue - 60.0) < 0.01);
// 50) 가용이 아닌 유닛: 가용 0, 몫 0, 용량 0
astAvail[1].bAvail := FALSE;
fbUv(iq_astView := astView, iq_astUnit := astUnit, iq_astAvail := astAvail, iq_astUnitCfg := astCfg,
	iq_astUnitEnv := astEnv, iq_astBatGroup := astBat, iq_astBatEnv := astBatEnv);
fbTally.M_Check(i_nId := 50, i_bOk := fbUv.q_astView[1].stView.nUnitAvail = 0 AND fbUv.q_astView[1].fRatingShare = 0.0 AND fbUv.q_astView[1].stView.fCapacity = 0.0
	AND ABS(fbUv.q_astView[1].stView.fPOut - 100.0) < 0.01);
astAvail[1].bAvail := TRUE;
END_ACTION

ACTION A_StdScheduleTest:
// 스탠다드 스케줄: EMS가 9시 방전 100, 10시 정지를 보내는 흐름 (한 스캔씩 직접 부름)
stStdView.stGroup.nUnitAvail := 1;
// 켜지기 전에 온 지령(번호 5, 50 kW)은 쓰지 않음
fbStd.i_astCmd[1].bUse		:= TRUE;	// [16번 수정 2026-11-09: 모드가 유닛마다 칸을 받음 (유닛 1 칸으로 시험). 원래 fbStd.i_stCmd, 출력 stStdOut.bPSetActive·fPSet]
fbStd.i_astCmd[1].bAlive	:= TRUE;
fbStd.i_astCmd[1].nPSeq		:= 5;
fbStd.i_astCmd[1].fP		:= 50.0;
fbStd.i_astCmd[1].nStateSeq	:= 3;
fbStd.i_astCmd[1].eState	:= E_PcsCmd.Run;
fbStd.M_Enter(i_stView := stStdView);
stStdOut := fbStd.M_Calc(i_stView := stStdView);
fbTally.M_Check(i_nId := 51, i_bOk := stStdOut.bUnitOut AND stStdOut.astUnit[1].bPSetActive AND stStdOut.astUnit[1].fPSet = 0.0 AND fbStd.q_nState = 3 AND NOT fbStd.q_abHold[1]);
// 9시: 방전 100 → 100, 다음 지령까지 유지
fbStd.i_astCmd[1].nPSeq	:= 6;
fbStd.i_astCmd[1].fP	:= 100.0;
stStdOut := fbStd.M_Calc(i_stView := stStdView);
stStdOut := fbStd.M_Calc(i_stView := stStdView);
fbTally.M_Check(i_nId := 52, i_bOk := ABS(stStdOut.astUnit[1].fPSet - 100.0) < 0.01 AND fbStd.q_nState = 0 AND fbStd.q_nCmdCount = 1);
// 10시: 정지 → 0 (새 P 지령 대기)
fbStd.i_astCmd[1].nStateSeq	:= 4;
fbStd.i_astCmd[1].eState	:= E_PcsCmd.Stop;
stStdOut := fbStd.M_Calc(i_stView := stStdView);
fbTally.M_Check(i_nId := 53, i_bOk := stStdOut.astUnit[1].bPSetActive AND stStdOut.astUnit[1].fPSet = 0.0 AND fbStd.q_nState = 3);
// Run만 다시 와도 옛 100은 되살아나지 않음
fbStd.i_astCmd[1].nStateSeq	:= 5;
fbStd.i_astCmd[1].eState	:= E_PcsCmd.Run;
stStdOut := fbStd.M_Calc(i_stView := stStdView);
fbTally.M_Check(i_nId := 54, i_bOk := stStdOut.astUnit[1].fPSet = 0.0 AND NOT fbStd.q_abHold[1]);
// 충전 -200 → -200. 이상값(무한대)은 버리고 앞 값 유지
fbStd.i_astCmd[1].nPSeq	:= 7;
fbStd.i_astCmd[1].fP	:= -200.0;
stStdOut := fbStd.M_Calc(i_stView := stStdView);
nBad0 := fbStd.q_nBadCount;
fbStd.i_astCmd[1].nPSeq	:= 8;
MEMCPY(destAddr := ADR(fInf), srcAddr := ADR(nInfBits), n := SIZEOF(fInf));	// +무한대 (비트로 만듦)
fbStd.i_astCmd[1].fP	:= fInf;
stStdOut := fbStd.M_Calc(i_stView := stStdView);
fbTally.M_Check(i_nId := 55, i_bOk := ABS(stStdOut.astUnit[1].fPSet + 200.0) < 0.01 AND fbStd.q_nBadCount = nBad0 + 1);
// EMS 끊김 → 0, 돌아와도 옛 값은 되살아나지 않음
fbStd.i_astCmd[1].bAlive := FALSE;
stStdOut := fbStd.M_Calc(i_stView := stStdView);
fbTally.M_Check(i_nId := 56, i_bOk := stStdOut.astUnit[1].fPSet = 0.0 AND fbStd.q_nState = 2);
fbStd.i_astCmd[1].bAlive := TRUE;
stStdOut := fbStd.M_Calc(i_stView := stStdView);
fbTally.M_Check(i_nId := 57, i_bOk := stStdOut.astUnit[1].fPSet = 0.0 AND fbStd.q_nState = 3);
fbStd.M_Exit();
END_ACTION

ACTION A_NanTest:
// NaN·무한대: 비트로 먼저 거르는지 (거르지 못하면 여기서 PLC가 멈춤)
MEMCPY(destAddr := ADR(fNan), srcAddr := ADR(nNanBits), n := SIZEOF(fNan));
// 58) F_IsFinite: NaN·무한대 FALSE, 보통 숫자 TRUE
fbTally.M_Check(i_nId := 58, i_bOk := NOT F_IsFinite(fNan) AND NOT F_IsFinite(fInf) AND F_IsFinite(-123.4) AND F_IsFinite(0.0));
// 59) F_CmdOk: NaN은 한도가 있든 없든 FALSE, 보통 숫자는 한도대로
fbTally.M_Check(i_nId := 59, i_bOk := NOT F_CmdOk(fNan, 0.0) AND NOT F_CmdOk(fNan, 1000.0) AND NOT F_CmdOk(fInf, 0.0)
	AND F_CmdOk(500.0, 1000.0) AND NOT F_CmdOk(1500.0, 1000.0));
// 60) 스탠다드 스케줄 모드: NaN P 지령은 버리고 앞 값 유지
fbStd.i_astCmd[1].bAlive	:= TRUE;
fbStd.M_Enter(i_stView := stStdView);
fbStd.i_astCmd[1].nPSeq		:= fbStd.i_astCmd[1].nPSeq + 1;
fbStd.i_astCmd[1].fP		:= 70.0;
stStdOut := fbStd.M_Calc(i_stView := stStdView);
nBad0 := fbStd.q_nBadCount;
fbStd.i_astCmd[1].nPSeq		:= fbStd.i_astCmd[1].nPSeq + 1;
fbStd.i_astCmd[1].fP		:= fNan;
stStdOut := fbStd.M_Calc(i_stView := stStdView);
fbTally.M_Check(i_nId := 60, i_bOk := ABS(stStdOut.astUnit[1].fPSet - 70.0) < 0.01 AND fbStd.q_nBadCount = nBad0 + 1);
fbStd.M_Exit();
// 61) EMS 명령 핸들러: 방전 NaN → 버리고 셈, P 번호 안 바뀜 (PCS1 = 칸 0)
nPSeq0 := fbEmsCmd.q_stCmd.anPcsPSeq[1];
nBad0 := fbEmsCmd.q_nBadValueCount;
astPcsRx[0].Value		:= fNan;
astPcsRx[0].CommandType	:= 5;
fbEmsCmd(i_nRxCount := 1, iq_astPcsCommand := astPcsRx, iq_astBatCommand := astBatRx);
fbTally.M_Check(i_nId := 61, i_bOk := fbEmsCmd.q_nBadValueCount = nBad0 + 1 AND fbEmsCmd.q_stCmd.anPcsPSeq[1] = nPSeq0 AND astPcsRx[0].CommandType = 0);
// 62) 상태 명령(Run)에 Value가 NaN이어도 명령은 받음 (값은 안 봄)
nRunSeq0 := fbEmsCmd.q_stCmd.astPcs[1].nSeq;
astPcsRx[0].Value		:= fNan;
astPcsRx[0].CommandType	:= 1;
fbEmsCmd(i_nRxCount := 2, iq_astPcsCommand := astPcsRx, iq_astBatCommand := astBatRx);
fbTally.M_Check(i_nId := 62, i_bOk := fbEmsCmd.q_stCmd.astPcs[1].nSeq = nRunSeq0 + 1 AND fbEmsCmd.q_stCmd.astPcs[1].eCmd = E_PcsCmd.Run);
// 63) 보통 값(방전 120)은 받음
astPcsRx[0].Value		:= 120.0;
astPcsRx[0].CommandType	:= 5;
fbEmsCmd(i_nRxCount := 3, iq_astPcsCommand := astPcsRx, iq_astBatCommand := astBatRx);
fbTally.M_Check(i_nId := 63, i_bOk := fbEmsCmd.q_stCmd.anPcsPSeq[1] = nPSeq0 + 1 AND ABS(fbEmsCmd.q_stCmd.afPcsP[1] - 120.0) < 0.01);
END_ACTION

END_PROGRAM

// ---- 20_Module/ControlMode/FB_CmStdSchedule.TcPOU
FUNCTION_BLOCK FB_CmStdSchedule EXTENDS FB_CtrlModeBase		// 제어 모드: 스탠다드 스케줄. 시간표를 PMS에 두지 않고 EMS가 시각마다 보내는 지령을 그대로 따름
// 예) 09~10시 방전 100 kW: EMS가 9시에 방전 100 kW, 10시에 정지를 보냄 → 이 모드는 받은 P를 다음 지령까지 유지하고, 정지 쪽 명령이 오면 버림
// Manual 지령과 같은 구조: 새 지령(번호가 바뀜)만 받음, 받은 값은 다음 지령까지 유지, 정지 쪽 명령 뒤에는 새 P 지령이 올 때까지 0
//   - 모드가 켜지기 전에 온 지령은 쓰지 않음 (켜진 뒤 새 지령부터). 켜져 있는 동안 P는 늘 냄 (지령이 없으면 0 → 등급이 낮은 다른 지령원 값이 새지 않게)
//   - EMS가 끊기면 받아 둔 P를 버리고 0. 이상값(NaN·무한대)은 버리고 앞 값을 유지 (정격 대비 상한은 코어 명령 필터)
//   - 상태 명령(Run·Stop 등) 자체는 EMS 지령원(FB_SrcEms)이 장비에 냄. 이 모드는 P만 냄. 역송 방지·방전 허용 시간은 걸지 않음 (EMS 책임, 코어 접속점 제한은 그대로)
// [16번 수정 2026-11-09: 유닛마다 따로 받고 유닛별 값(bUnitOut)으로 냄. 제어 모드 관리자가 접속점 그룹 단위여도 EMS가 PCS마다 보낸 값을 그대로 따름.
//   원래는 PCS마다 관리자·모드 인스턴스(g_fbCmStdSched1·2)가 있고 지령 하나(i_stCmd)를 그 관리자 단위 값으로 냄]
// 입력 i_astCmd는 MAIN(A_PassEmsCmd)이 매 스캔 채움 (PCS 지령을 그 PCS의 유닛에 정격 비율로 나눔)
VAR_INPUT
	i_astCmd	: ARRAY[1..GVL_PARAM.UNIT_COUNT] OF ST_CmExtCmd;	// 유닛마다 바깥 지령. bUse FALSE인 칸은 내지 않음
END_VAR
VAR_OUTPUT
	q_nState	: UINT;				// 요약: 0 = 쓰는 유닛 모두 받은 P를 냄, 그 외 = 0을 내는 유닛의 첫 이유 (M_ReasonText)
	q_anState	: ARRAY[1..GVL_PARAM.UNIT_COUNT] OF UINT;	// 유닛마다 0 = 받은 P를 냄, 그 외 = 0을 내는 이유
	q_abHold	: ARRAY[1..GVL_PARAM.UNIT_COUNT] OF BOOL;	// 받아 둔 P 지령 있음
	q_afPCmd	: ARRAY[1..GVL_PARAM.UNIT_COUNT] OF REAL;	// kW, 받아 둔 P 지령 (q_abHold일 때)
	q_nCmdCount	: UDINT;			// 켜진 뒤 받은 P 지령 수 (유닛 합)
	q_nBadCount	: UDINT;			// 이상값이라 버린 P 지령 수
END_VAR
VAR
	_anPSeq		: ARRAY[1..GVL_PARAM.UNIT_COUNT] OF UDINT;	// 처리한 P 지령 번호
	_anStateSeq	: ARRAY[1..GVL_PARAM.UNIT_COUNT] OF UDINT;	// 처리한 상태 명령 번호
END_VAR
VAR CONSTANT
	RSN_NO_UNIT		: UINT := 1;	// 진입 거부: 가용 유닛 없음
	RSN_NO_EXT		: UINT := 2;	// EMS 끊김 → 0
	RSN_WAIT_CMD	: UINT := 3;	// 새 P 지령 대기 (켜진 뒤 아직 없음, 또는 정지 쪽 명령 뒤) → 0
END_VAR

METHOD M_CheckEnter : UINT
VAR_INPUT
	i_stView	: ST_CtrlModeView;	// 그룹 값(stGroup)·현지 시각(stTime). 관리자가 매 스캔 채움
END_VAR
M_CheckEnter := 0;
IF i_stView.stGroup.nUnitAvail = 0 THEN
	M_CheckEnter := RSN_NO_UNIT;
END_IF
END_METHOD

METHOD M_Enter
VAR_INPUT
	i_stView	: ST_CtrlModeView;	// 그룹 값(stGroup)·현지 시각(stTime). 관리자가 매 스캔 채움
END_VAR
VAR
	u			: UINT;
END_VAR
SUPER^.M_Enter(i_stView := i_stView);
// 켜지기 전에 온 지령은 쓰지 않음: 지금 번호를 처리한 것으로 두고 새 지령을 기다림
FOR u := 1 TO GVL_PARAM.UNIT_COUNT DO
	_anPSeq[u]		:= i_astCmd[u].nPSeq;
	_anStateSeq[u]	:= i_astCmd[u].nStateSeq;
	q_abHold[u]		:= FALSE;
	q_afPCmd[u]		:= 0.0;
END_FOR
q_nCmdCount	:= 0;
END_METHOD

METHOD M_Calc : ST_CtrlModeOut
VAR_INPUT
	i_stView	: ST_CtrlModeView;	// 그룹 값(stGroup)·현지 시각(stTime). 관리자가 매 스캔 채움
END_VAR
VAR
	u			: UINT;
	bNewCmd		: BOOL;		// 이번 스캔에 새 지령이 옴 (살아 있다는 표시)
	bAlive		: BOOL;
END_VAR
q_nState := 0;
FOR u := 1 TO GVL_PARAM.UNIT_COUNT DO
	bNewCmd := i_astCmd[u].nStateSeq <> _anStateSeq[u] OR i_astCmd[u].nPSeq <> _anPSeq[u];
	// 1) 상태 명령: 정지 쪽이면 받아 둔 P를 버림 (같은 메시지에 P가 같이 오면 아래에서 P가 다시 들어감)
	IF i_astCmd[u].nStateSeq <> _anStateSeq[u] THEN
		_anStateSeq[u] := i_astCmd[u].nStateSeq;
		IF i_astCmd[u].eState = E_PcsCmd.Stop OR i_astCmd[u].eState = E_PcsCmd.Standby OR i_astCmd[u].eState = E_PcsCmd.EStop THEN
			q_abHold[u] := FALSE;
		END_IF
	END_IF
	// 2) 새 P 지령: 다음 지령까지 유지. 이상값은 버리고 앞 값 유지
	IF i_astCmd[u].nPSeq <> _anPSeq[u] THEN
		_anPSeq[u] := i_astCmd[u].nPSeq;
		IF F_CmdOk(i_fValue := i_astCmd[u].fP, i_fLimit := 0.0) THEN
			q_abHold[u]	:= TRUE;
			q_afPCmd[u]	:= i_astCmd[u].fP;
			q_nCmdCount	:= q_nCmdCount + 1;
		ELSE
			q_nBadCount	:= q_nBadCount + 1;
		END_IF
	END_IF
	// 3) EMS가 끊기면 버림 (돌아와도 옛 지령이 되살아나지 않음).
	//    bAlive는 지난 스캔 값이라, 조용하던 EMS의 첫 지령 스캔에는 아직 FALSE → 새 지령이 온 스캔은 살아 있는 것으로 봄
	bAlive := i_astCmd[u].bAlive OR bNewCmd;
	IF NOT bAlive THEN
		q_abHold[u] := FALSE;
	END_IF
	// 4) 유닛 상태·출력: 쓰는 유닛은 켜져 있는 동안 P를 늘 냄. Q는 다른 지령원에 맡김
	IF q_abHold[u] THEN
		q_anState[u] := 0;
	ELSIF NOT bAlive THEN
		q_anState[u] := RSN_NO_EXT;
	ELSE
		q_anState[u] := RSN_WAIT_CMD;
	END_IF
	M_Calc.astUnit[u].bPSetActive	:= i_astCmd[u].bUse;
	M_Calc.astUnit[u].fPSet			:= SEL(q_abHold[u], 0.0, q_afPCmd[u]);
	M_Calc.astUnit[u].bQSetActive	:= FALSE;
	M_Calc.astUnit[u].fQSet			:= 0.0;
	IF i_astCmd[u].bUse AND q_nState = 0 THEN
		q_nState := q_anState[u];
	END_IF
END_FOR
M_Calc.bUnitOut		:= TRUE;		// 접속점 그룹 값(bPSetActive·fPSet)은 쓰지 않음
M_Calc.bPSetActive	:= FALSE;
M_Calc.fPSet		:= 0.0;
M_Calc.bQSetActive	:= FALSE;
M_Calc.fQSet		:= 0.0;
M_Calc.bExitReq		:= FALSE;
M_Calc.nReason		:= q_nState;
END_METHOD

METHOD M_ReasonText : WSTRING(63)
VAR_INPUT
	i_nReason	: UINT;
END_VAR
CASE i_nReason OF
	RSN_NO_UNIT:	M_ReasonText := "스탠다드 스케줄: 가용 유닛 없음";
	RSN_NO_EXT:		M_ReasonText := "스탠다드 스케줄: EMS 끊김 (0)";
	RSN_WAIT_CMD:	M_ReasonText := "스탠다드 스케줄: 새 P 지령 대기 (0)";
ELSE
	M_ReasonText := WCONCAT("이유 ", TO_WSTRING(i_nReason));
END_CASE
END_METHOD

END_FUNCTION_BLOCK

// ---- 99_Test/PRG_TestStdLive.TcPOU
PROGRAM PRG_TestStdLive		// 스탠다드 스케줄 모드 실제 경로 시험 (시험 모드, MAIN이 부름): EMS 명령 레코드 → FB_EmsCommand(MqttTask) → GVL_IF → MAIN A_PassEmsCmd → 모드 → 관리자 → 코어 고르기
// bStart := TRUE로 시작. PCS2(유닛 2)를 Auto로 두고 접속점 그룹 관리자(g_fbCtrlMode1)에 모드 5 (유닛 2 칸을 봄).
// [16번 수정 2026-11-09: 관리자 2(g_fbCtrlMode2)·모드 g_fbCmStdSched2 → 접속점 그룹 관리자 g_fbCtrlMode1·g_fbCmStdSched1의 유닛 2 칸] EMS 명령은 MQTT 수신 칸(GVL_MQTT.g_astPcsCommand[1] = PCS2)에 직접 넣음 (브로커 없이)
// A: 켠 직후 EMS P 없음 → 0 / B: 방전 100 → 100 / C: 충전 50 → -50 / D: 정지 → 0 (새 P 지령 대기)
// 조건이 2 s 이어지면 통과. 장비 쓰기(DEVICE_WRITE)와 무관하게 코어 고르기 결과(MAIN.fbSelect)까지 봄. 끝나면 모드 0, 운전 모드를 되돌림
VAR
	bStart		: BOOL;
	bDone		: BOOL;
	bPass		: BOOL;
	nStep		: UINT;
	wsStep		: WSTRING(80);
	wsFail		: WSTRING(80);
	(* 지금 값 *)
	nActive		: UINT;			// 접속점 그룹 관리자 켜진 모드 (5 = 스탠다드 스케줄)
	nModeState	: UINT;			// 모드 q_nState (0 = P 냄, 2 = EMS 끊김, 3 = 새 지령 대기)
	fModeP		: REAL;			// 모드가 받아 둔 P
	bEmsAlive	: BOOL;			// EMS 지령원 유효
	fMgrP		: REAL;			// 접속점 그룹 관리자 출력 (유닛 2 칸)
	bMgrP		: BOOL;
	stPick		: ST_Pick;		// 코어 고르기 결과 (Auto 유닛 2)
	(* 판정 *)
	bA			: BOOL;
	bB			: BOOL;
	bC			: BOOL;
	bD			: BOOL;
	fB			: REAL;
	fC			: REAL;
	(* 내부 *)
	nU2			: UINT := 2;
	eOpModeBak	: E_OpMode;
	bBackedUp	: BOOL;
	bCond		: BOOL;
	nLastStep	: UINT;
	tonStep		: TON;
	tonOk		: TON;
	stOut		: ST_SourceOutput;
END_VAR

// 지금 값
nActive		:= GVL_SITE.g_fbCtrlMode1.q_nActive;
stOut		:= GVL_SITE.g_fbCtrlMode1.Output;
IF nU2 >= 1 AND nU2 <= GVL_PARAM.UNIT_COUNT THEN
	nModeState	:= GVL_SITE.g_fbCmStdSched1.q_anState[nU2];
	fModeP		:= GVL_SITE.g_fbCmStdSched1.q_afPCmd[nU2];
	bEmsAlive	:= GVL_SITE.g_fbCmStdSched1.i_astCmd[nU2].bAlive;
	bMgrP	:= stOut.astUnit[nU2].bPSetActive;
	fMgrP	:= stOut.astUnit[nU2].fPSet;
	stPick	:= MAIN.fbSelect.q_astAutoUnitP[nU2];
END_IF

tonStep(IN := nStep >= 20 AND nStep < 900, PT := T#30S);
bCond := FALSE;

CASE nStep OF
	0:
		IF bStart THEN
			bStart := FALSE;	bDone := FALSE;	bPass := FALSE;	wsFail := "";
			bA := FALSE;	bB := FALSE;	bC := FALSE;	bD := FALSE;
			nStep := 10;
		ELSIF NOT bDone THEN
			wsStep := "대기: bStart := TRUE로 시작";
		END_IF

	10:	// PCS2 Auto
		wsStep := "PCS2 Auto 전환";
		IF nU2 > GVL_PARAM.UNIT_COUNT OR GVL_PARAM.PCS_COUNT < 2 THEN
			wsFail := "PCS·유닛이 2개 이상이어야 함";
			nStep := 900;
		ELSE
			eOpModeBak	:= GVL_PERSIST.g_aeOpMode[nU2];
			bBackedUp	:= TRUE;
			GVL_PERSIST.g_aeOpMode[nU2] := E_OpMode.Auto;
			nStep := 20;
		END_IF

	20:
		wsStep := "Auto 전환 대기";
		IF MAIN.fbModeSwitch.q_aeOpMode[nU2] = E_OpMode.Auto THEN
			GVL_SITE.g_fbCtrlMode1.i_nModeReq := 5;
			GVL_SITE.g_fbCtrlMode1.i_bRetry := TRUE;
			nStep := 30;
		END_IF

	30:
		wsStep := "스탠다드 스케줄 모드 켜는 중";
		IF nActive = 5 THEN
			nStep := 100;
		ELSIF GVL_SITE.g_fbCtrlMode1.q_eRefuse <> E_CtrlModeRefuse.None THEN
			wsFail := WCONCAT("모드 거부: ", GVL_SITE.g_fbCtrlMode1.M_ModeReasonText(i_nSlot := 5, i_nReason := GVL_SITE.g_fbCtrlMode1.q_nRefuseReason));
			nStep := 900;
		END_IF

	100: // A: 켠 직후, EMS P 없음 → 0
		wsStep := "A: EMS P 없음 → 0";
		bCond := nActive = 5 AND (nModeState = 3 OR nModeState = 2) AND bMgrP AND fMgrP = 0.0;
		IF tonOk.Q THEN
			bA := TRUE;
			M_Send(i_nType := 5, i_fValue := 100.0);		// 방전 100
			nStep := 110;
		END_IF
	110: // B: 방전 100
		wsStep := "B: EMS 방전 100 → 100";
		bCond := nModeState = 0 AND ABS(fModeP - 100.0) < 0.01 AND bMgrP AND ABS(fMgrP - 100.0) < 0.01
			AND stPick.bActive AND ABS(stPick.fValue - 100.0) < 0.01 AND stPick.nModule = GVL_SITE.g_fbCtrlMode1.ModuleId;
		IF tonOk.Q THEN
			bB := TRUE;	fB := stPick.fValue;
			M_Send(i_nType := 4, i_fValue := 50.0);		// 충전 50
			nStep := 120;
		END_IF
	120: // C: 충전 50
		wsStep := "C: EMS 충전 50 → -50";
		bCond := nModeState = 0 AND ABS(fMgrP + 50.0) < 0.01 AND stPick.bActive AND ABS(stPick.fValue + 50.0) < 0.01;
		IF tonOk.Q THEN
			bC := TRUE;	fC := stPick.fValue;
			M_Send(i_nType := 2, i_fValue := 0.0);		// 정지
			nStep := 130;
		END_IF
	130: // D: 정지 → 0 (새 P 지령 대기)
		wsStep := "D: EMS 정지 → 0";
		bCond := nModeState = 3 AND bMgrP AND fMgrP = 0.0 AND stPick.bActive AND stPick.fValue = 0.0;
		IF tonOk.Q THEN
			bD := TRUE;
			nStep := 900;
		END_IF

	900: // 정리
		GVL_SITE.g_fbCtrlMode1.i_nModeReq := 0;
		IF bBackedUp THEN
			GVL_PERSIST.g_aeOpMode[nU2] := eOpModeBak;
			bBackedUp := FALSE;
		END_IF
		bPass := bA AND bB AND bC AND bD AND wsFail = "";
		bDone := TRUE;
		IF bPass THEN
			wsStep := "끝: 통과";
		ELSE
			wsStep := "끝: 실패 (wsFail·구간 결과 확인)";
		END_IF
		nStep := 0;
END_CASE

tonOk(IN := bCond AND nStep = nLastStep, PT := T#2S);
IF tonStep.Q AND nStep >= 20 AND nStep < 900 THEN
	wsFail	:= WCONCAT("시간 초과: ", wsStep);
	nStep	:= 900;
END_IF
IF nStep <> nLastStep THEN
	tonStep(IN := FALSE);
	tonOk(IN := FALSE);
	nLastStep := nStep;
END_IF

METHOD PRIVATE M_Send		// EMS 명령 레코드 하나를 MQTT 수신 칸에 넣음 (PCS2 = 칸 1). 값을 먼저, 종류를 마지막에 (MqttTask가 종류를 보고 처리)
VAR_INPUT
	i_nType		: UDINT;	// PCS CommandType: 1 Run, 2 Stop, 3 Standby, 4 충전, 5 방전
	i_fValue	: REAL;		// kW
END_VAR
GVL_MQTT.g_astPcsCommand[1].DeviceIndex	:= 2;	// PCS2 (번호 1부터) [1부터 2026-11-10]
GVL_MQTT.g_astPcsCommand[1].Value		:= i_fValue;
GVL_MQTT.g_astPcsCommand[1].CommandType	:= i_nType;
END_METHOD

END_PROGRAM

// ---- 90_Project/PRG_Redundancy.TcPOU
PROGRAM PRG_Redundancy		// 이중화 태스크에서 부름 (높은 우선순위). 이 PLC의 역할(Primary/Secondary)과 지금 장비에 쓰는지(Active)를 GVL_IF에 씀
VAR
	fbGetNetId		: FB_GetLocalAmsNetID;	// 이 PLC의 AMS Net ID 읽기 (시작 때 한 번)
	sMyNetId		: T_AmsNetId;			// 읽은 이 PLC의 Net ID (온라인 확인용: RED_SET에 적을 값)
	bNetIdRead		: BOOL;					// Net ID를 읽었음
	tLastScan		: TIME;				// 지난 스캔의 시스템 시각 (멈췄다 이어짐 감지)
	bScanned		: BOOL;				// 첫 스캔을 지남 (시작 때는 이어짐으로 안 봄)
	bResume			: BOOL;				// 이번 스캔이 멈췄다 이어진 첫 스캔
	fbRedSync		: FB_RedSync;			// 운영 설정 동기화 (Active → Standby)
	fbRedState		: FB_RedState;			// 역할 + 상대 상태 → Active 판단
	fbRedLink		: FB_RedLink;			// 상대 PLC와 EAP 하트비트·접점 신호 (I/O는 이 인스턴스에 연결)
END_VAR

(* 0) 멈췄다 이어짐 감지: ADS·XAE의 Stop/Run은 변수를 초기화하지 않고 이어서 돎. 이전 스캔과 시스템 시각이 1 s 넘게 벌어지면 멈췄던 것으로 보고 상태를 Init부터 다시 정함 *)
bResume := bScanned AND (TIME() - tLastScan) > T#1S;
bScanned := TRUE;
tLastScan := TIME();
IF bResume AND GVL_SITE.RED_SET.bUse THEN
	GVL_IF.g_nRedResumeCount	:= GVL_IF.g_nRedResumeCount + 1;
	GVL_IF.g_bRedActive			:= FALSE;		// 옛 Active를 상대에게 알리거나 장비에 쓰지 않도록 이 스캔부터 내림
	GVL_IF.g_bRedWrite			:= FALSE;
	GVL_IF.g_eRedState			:= E_RedState.Init;
END_IF

(* 1) 역할: 이중화를 안 쓰면 Primary. 쓰면 이 PLC Net ID를 GVL_SITE.RED_SET과 비교 *)
IF NOT GVL_SITE.RED_SET.bUse THEN
	GVL_IF.g_eRedRole := E_RedRole.Primary;
ELSIF NOT bNetIdRead THEN
	GVL_IF.g_eRedRole := E_RedRole.Reading;
	fbGetNetId(bExecute := TRUE);
	IF NOT fbGetNetId.bBusy THEN
		IF NOT fbGetNetId.bError THEN
			sMyNetId	:= fbGetNetId.AddrString;
			bNetIdRead	:= TRUE;
		END_IF
		fbGetNetId(bExecute := FALSE);		// 오류면 다음 스캔에 다시 읽음
	END_IF
ELSIF sMyNetId = GVL_SITE.RED_SET.sPrimaryNetId THEN
	GVL_IF.g_eRedRole := E_RedRole.Primary;
ELSIF sMyNetId = GVL_SITE.RED_SET.sSecondaryNetId THEN
	GVL_IF.g_eRedRole := E_RedRole.Secondary;
ELSE
	GVL_IF.g_eRedRole := E_RedRole.NoMatch;		// 설정 오류 (FB_ConfigCheck)
END_IF

(* 2) 상대 PLC 상태: EAP 하트비트와 접점 신호를 보고 판정. 이중화를 안 쓰면 보내지도 않음. 내 Active는 지난 스캔 값을 보냄 *)
IF GVL_SITE.RED_SET.bUse THEN
	fbRedLink(	i_stSet	:= GVL_SITE.RED_SET,
				i_eRole	:= GVL_IF.g_eRedRole,
				i_bActive	:= GVL_IF.g_bRedActive,
				i_eState	:= GVL_IF.g_eRedState);
	GVL_IF.g_nRedSeq			:= fbRedLink.q_nTxCount;
	GVL_IF.g_ePeerState		:= fbRedLink.q_ePeer;
	GVL_IF.g_bPeerEapOk		:= fbRedLink.q_bEapOk;
	GVL_IF.g_bPeerWireOk		:= fbRedLink.q_bWireOk;
	GVL_IF.g_nPeerRole		:= fbRedLink.q_stPeer.nRole;
	GVL_IF.g_bPeerActive		:= fbRedLink.q_stPeer.bActive;
	GVL_IF.g_nPeerState		:= fbRedLink.q_stPeer.nState;
	GVL_IF.g_bPeerWireActive	:= fbRedLink.q_bPeerWireActive;
	GVL_IF.g_bRedRoleConflict	:= fbRedLink.q_bRoleConflict;
ELSE
	GVL_IF.g_ePeerState		:= E_RedPeer.Unknown;
	GVL_IF.g_bPeerEapOk		:= FALSE;
	GVL_IF.g_bPeerWireOk		:= FALSE;
	GVL_IF.g_bRedRoleConflict	:= FALSE;
	GVL_IF.g_nPeerState		:= 0;
END_IF

(* 3) 동기화: 운영 설정을 상대에게 보내고, 내가 Active가 아니고 상대가 Active이면 받은 값으로 맞춤
   동기화 대상 = GVL_PERSIST의 운영 설정 (재기동 기록·모듈 설정 묶음 제외) + 제어 모드 요청. 대상을 늘리면 ST_RedSyncCfg와 FB_RedSync의 보내기·맞추기에 추가 *)
IF GVL_SITE.RED_SET.bUse THEN
	fbRedSync(	i_bUse		:= TRUE,
				i_bApply	:= GVL_IF.g_eRedState <> E_RedState.Active AND GVL_IF.g_bPeerEapOk AND GVL_IF.g_bPeerActive);
	GVL_IF.g_bSyncInSync	:= fbRedSync.q_bInSync;
	GVL_IF.g_bSyncFresh		:= fbRedSync.q_bFresh;
	GVL_IF.g_nSyncApplied	:= fbRedSync.q_nApplied;
ELSE
	GVL_IF.g_bSyncInSync	:= FALSE;
	GVL_IF.g_bSyncFresh		:= FALSE;
END_IF

(* 4) Active: 역할과 상대 상태로 정함 (FB_RedState). 두 PLC가 동시에 Active가 되지 않음. Secondary 승격(절체)·Primary 복귀 포함 *)
fbRedState(	i_bUse			:= GVL_SITE.RED_SET.bUse,
			i_stSet			:= GVL_SITE.RED_SET,
			i_eRole			:= GVL_IF.g_eRedRole,
			i_ePeer			:= GVL_IF.g_ePeerState,
			i_bPeerActive	:= (GVL_IF.g_bPeerEapOk AND GVL_IF.g_bPeerActive) OR (GVL_IF.g_bPeerWireOk AND GVL_IF.g_bPeerWireActive),
			i_bPeerHandover	:= GVL_IF.g_bPeerEapOk AND GVL_IF.g_nPeerState = TO_INT(E_RedState.Handover),
			i_bRoleConflict	:= GVL_IF.g_bRedRoleConflict,
			i_bReset		:= bResume AND GVL_SITE.RED_SET.bUse,
			i_bSyncDone		:= GVL_IF.g_bSyncInSync);
GVL_IF.g_eRedState	:= fbRedState.q_eState;
GVL_IF.g_bRedActive	:= fbRedState.q_bActive;
GVL_IF.g_bRedWrite	:= fbRedState.q_bWrite;
GVL_IF.g_nRedSwitchCount	:= fbRedState.q_nSwitchCount;
GVL_IF.g_eRedSwitch	:= fbRedState.q_eLastSwitch;

END_PROGRAM

